(* IEC 61131-3 sources: plc-process-lib/tests/POUs/Suites/FB_Pid_Test, 85 files *)

(* ---- AntiWindupLongSaturationRecoversWithinTt.method.decl.st ---- *)
// Anti-windup обратным расчётом (Kp = 1, Ti = 10 с, Tt = авто = Ti): 60 с на верхнем пределе при
// ошибке +20 %, затем ошибка -20 %. С обратным расчётом интегратор ограничен (v ≈ 100 + Tt·Kp·e/Ti)
// и выход уходит с предела сразу; для сравнения тот же ФБ с Tt = 1·10^6 с (обратного расчёта
// практически нет) остаётся на пределе и через Tt после смены знака.
METHOD PRIVATE AntiWindupLongSaturationRecoversWithinTt
VAR
    fbTime    : FB_FakeTime;       // подменное время, старт 1 ч
    fbPidAw   : FB_PID;            // ФБ под тестом: Tt = авто
    fbPidNoAw : FB_PID;            // сравнение: Tt = 1e6 с
    stCmdAw   : ST_PidCmd;         // команды
    stCmdNoAw : ST_PidCmd;
    stRetAw   : ST_DeviceRetain;   // режим: старт в Manual
    stRetNoAw : ST_DeviceRetain;
    stCfgAw   : ST_PidCfg;         // конфигурация
    stCfgNoAw : ST_PidCfg;
    iStep     : INT;               // шаг цикла
    rOutSatAw : REAL;              // выход в конце насыщения
    rISatAw   : REAL;              // интегратор в конце насыщения
    rISatNoAw : REAL;
    rOutRevAw : REAL;              // выход в первом шаге после смены знака ошибки
    rOutRevNo : REAL;
END_VAR

(* ---- AntiWindupLongSaturationRecoversWithinTt.method.impl.st ---- *)
coUnit.TEST('Pid_AntiWindup_LongSaturation_RecoversWithinTt');
// источник: tools/reference/pid.py, сценарий aw_recovery
stCfgAw.rKp := 1.0;
stCfgAw.rTi_s := 10.0;
stCfgAw.rTt_s := 0.0;
stCfgNoAw := stCfgAw;
stCfgNoAw.rTt_s := 1.0E6;
stCmdAw.rManualOut_pct := 50.0;
stCmdAw.rSp_eu := 50.0;
stCmdNoAw := stCmdAw;
fbPidAw.rPv_eu := 50.0;
fbPidAw.xPvValid := TRUE;
fbPidNoAw.rPv_eu := 50.0;
fbPidNoAw.xPvValid := TRUE;
fbPidAw(itfTime := fbTime, stCmd := stCmdAw, stRetain := stRetAw, stCfg := stCfgAw);          // t0: Manual
fbPidNoAw(itfTime := fbTime, stCmd := stCmdNoAw, stRetain := stRetNoAw, stCfg := stCfgNoAw);
fbTime.Advance(tStep := T#100MS);
stCmdAw.stCommon.xSetAuto := TRUE;
stCmdNoAw.stCommon.xSetAuto := TRUE;
fbPidAw(itfTime := fbTime, stCmd := stCmdAw, stRetain := stRetAw, stCfg := stCfgAw);          // Auto
fbPidNoAw(itfTime := fbTime, stCmd := stCmdNoAw, stRetain := stRetNoAw, stCfg := stCfgNoAw);
fbPidAw.rPv_eu := 30.0;                                                                         // e = +20 %
fbPidNoAw.rPv_eu := 30.0;
FOR iStep := 1 TO 600 DO                                                                        // 60 с
    fbTime.Advance(tStep := T#100MS);
    fbPidAw(itfTime := fbTime, stCmd := stCmdAw, stRetain := stRetAw, stCfg := stCfgAw);
    fbPidNoAw(itfTime := fbTime, stCmd := stCmdNoAw, stRetain := stRetNoAw, stCfg := stCfgNoAw);
END_FOR
rOutSatAw := fbPidAw.rOut_pct;
rISatAw := fbPidAw.stSts.rI_pct;
rISatNoAw := fbPidNoAw.stSts.rI_pct;
fbPidAw.rPv_eu := 70.0;                                                                         // e = -20 %
fbPidNoAw.rPv_eu := 70.0;
fbTime.Advance(tStep := T#100MS);
fbPidAw(itfTime := fbTime, stCmd := stCmdAw, stRetain := stRetAw, stCfg := stCfgAw);
fbPidNoAw(itfTime := fbTime, stCmd := stCmdNoAw, stRetain := stRetNoAw, stCfg := stCfgNoAw);
rOutRevAw := fbPidAw.rOut_pct;
rOutRevNo := fbPidNoAw.rOut_pct;
FOR iStep := 1 TO 99 DO                                                                         // до Tt = 10 с
    fbTime.Advance(tStep := T#100MS);
    fbPidAw(itfTime := fbTime, stCmd := stCmdAw, stRetain := stRetAw, stCfg := stCfgAw);
    fbPidNoAw(itfTime := fbTime, stCmd := stCmdNoAw, stRetain := stRetNoAw, stCfg := stCfgNoAw);
END_FOR
// ref: aw_recovery.out_sat_aw
AssertEquals_REAL(Expected := 100.0, Actual := rOutSatAw, Delta := 1.0E-4, Message := 'saturated at rOutMax_pct');
// ref: aw_recovery.i_sat_aw
AssertEquals_REAL(Expected := 99.782799, Actual := rISatAw, Delta := 1.0E-3,
                  Message := 'I bounded by back-calculation');
// ref: aw_recovery.i_sat_noaw
AssertEquals_REAL(Expected := 169.997986, Actual := rISatNoAw, Delta := 1.0E-3, Message := 'I winds up without it');
// ref: aw_recovery.out_rev_aw
AssertEquals_REAL(Expected := 79.782799, Actual := rOutRevAw, Delta := 1.0E-3, Message := 'leaves limit at once');
// ref: aw_recovery.out_rev_noaw
AssertEquals_REAL(Expected := 100.0, Actual := rOutRevNo, Delta := 1.0E-4, Message := 'wound-up: still at limit');
// ref: aw_recovery.out_tt_aw
AssertEquals_REAL(Expected := 59.982796, Actual := fbPidAw.rOut_pct, Delta := 1.0E-3, Message := 'recovered within Tt');
// ref: aw_recovery.out_tt_noaw
AssertEquals_REAL(Expected := 100.0, Actual := fbPidNoAw.rOut_pct, Delta := 1.0E-4, Message := 'wound-up after Tt');
AssertFalse(Condition := fbPidAw.xSatHigh, Message := 'back-calculation: not saturated after Tt');
coUnit.TEST_FINISHED();

(* ---- AntiWindupOutActFeedbackTracksExternalLimit.method.decl.st ---- *)
// Обратный расчёт по фактическому выходу (xUseOutAct): механизм не опускается ниже 30 % (минимум
// частоты ПЧ), rOutAct_pct = MAX(30, выход прошлого вызова). При ошибке -10 % 60 с выход ПИД
// держится у внешнего предела (около 30 - Tt·Kp·|e|/Ti = 20 %), а не уходит в 0; после смены
// знака ошибки механизм отвечает сразу. Без xUseOutAct ПИД уходит в 0 и после смены знака
// остаётся ниже 30 %.
METHOD PRIVATE AntiWindupOutActFeedbackTracksExternalLimit
VAR
    fbTime     : FB_FakeTime;       // подменное время, старт 1 ч
    fbPidAct   : FB_PID;            // ФБ под тестом: xUseOutAct
    fbPidNoAct : FB_PID;            // сравнение: без xUseOutAct
    stCmdAct   : ST_PidCmd;         // команды
    stCmdNoAct : ST_PidCmd;
    stRetAct   : ST_DeviceRetain;   // режим: старт в Manual
    stRetNoAct : ST_DeviceRetain;
    stCfgAct   : ST_PidCfg;         // конфигурация
    stCfgNoAct : ST_PidCfg;
    iStep      : INT;               // шаг цикла
    rHoldAct   : REAL;              // выход в конце 60 с
    rHoldNoAct : REAL;
END_VAR

(* ---- AntiWindupOutActFeedbackTracksExternalLimit.method.impl.st ---- *)
coUnit.TEST('Pid_AntiWindup_OutActFeedback_TracksExternalLimit');
// источник: tools/reference/pid.py, сценарий outact
stCfgAct.rKp := 1.0;
stCfgAct.rTi_s := 10.0;
stCfgNoAct := stCfgAct;
stCfgAct.xUseOutAct := TRUE;
stCmdAct.rManualOut_pct := 50.0;
stCmdAct.rSp_eu := 50.0;
stCmdNoAct := stCmdAct;
fbPidAct.rPv_eu := 50.0;
fbPidAct.xPvValid := TRUE;
fbPidNoAct.rPv_eu := 50.0;
fbPidNoAct.xPvValid := TRUE;
fbPidAct(itfTime := fbTime, stCmd := stCmdAct, stRetain := stRetAct, stCfg := stCfgAct);          // t0: Manual
fbPidNoAct(itfTime := fbTime, stCmd := stCmdNoAct, stRetain := stRetNoAct, stCfg := stCfgNoAct);
fbPidAct.rOutAct_pct := MAX(30.0, fbPidAct.rOut_pct);
fbPidNoAct.rOutAct_pct := MAX(30.0, fbPidNoAct.rOut_pct);
fbTime.Advance(tStep := T#100MS);
stCmdAct.stCommon.xSetAuto := TRUE;
stCmdNoAct.stCommon.xSetAuto := TRUE;
fbPidAct(itfTime := fbTime, stCmd := stCmdAct, stRetain := stRetAct, stCfg := stCfgAct);          // Auto
fbPidNoAct(itfTime := fbTime, stCmd := stCmdNoAct, stRetain := stRetNoAct, stCfg := stCfgNoAct);
fbPidAct.rPv_eu := 60.0;                                                                            // e = -10 %
fbPidNoAct.rPv_eu := 60.0;
FOR iStep := 1 TO 600 DO                                                                            // 60 с
    fbPidAct.rOutAct_pct := MAX(30.0, fbPidAct.rOut_pct);
    fbPidNoAct.rOutAct_pct := MAX(30.0, fbPidNoAct.rOut_pct);
    fbTime.Advance(tStep := T#100MS);
    fbPidAct(itfTime := fbTime, stCmd := stCmdAct, stRetain := stRetAct, stCfg := stCfgAct);
    fbPidNoAct(itfTime := fbTime, stCmd := stCmdNoAct, stRetain := stRetNoAct, stCfg := stCfgNoAct);
END_FOR
rHoldAct := fbPidAct.rOut_pct;
rHoldNoAct := fbPidNoAct.rOut_pct;
fbPidAct.rPv_eu := 40.0;                                                                            // e = +10 %
fbPidNoAct.rPv_eu := 40.0;
FOR iStep := 1 TO 30 DO                                                                             // 3 с
    fbPidAct.rOutAct_pct := MAX(30.0, fbPidAct.rOut_pct);
    fbPidNoAct.rOutAct_pct := MAX(30.0, fbPidNoAct.rOut_pct);
    fbTime.Advance(tStep := T#100MS);
    fbPidAct(itfTime := fbTime, stCmd := stCmdAct, stRetain := stRetAct, stCfg := stCfgAct);
    fbPidNoAct(itfTime := fbTime, stCmd := stCmdNoAct, stRetain := stRetNoAct, stCfg := stCfgNoAct);
END_FOR
// ref: outact.out_hold_act
AssertEquals_REAL(Expected := 20.067717, Actual := rHoldAct, Delta := 1.0E-3, Message := 'held near external limit');
// ref: outact.out_hold_noact
AssertEquals_REAL(Expected := 0.0, Actual := rHoldNoAct, Delta := 1.0E-4, Message := 'without OutAct: down to 0');
// ref: outact.out_rev_act
AssertEquals_REAL(Expected := 42.839634, Actual := fbPidAct.rOut_pct, Delta := 1.0E-3, Message := 'responds at once');
// ref: outact.out_rev_noact
AssertEquals_REAL(Expected := 14.239797, Actual := fbPidNoAct.rOut_pct, Delta := 1.0E-3, Message := 'still below 30 %');
AssertTrue(Condition := fbPidAct.rOut_pct > 30.0, Message := 'with OutAct the actuator moves above its minimum');
AssertTrue(Condition := fbPidNoAct.rOut_pct < 30.0, Message := 'without OutAct the actuator still sits at 30 %');
coUnit.TEST_FINISHED();

(* ---- AntiWindupOutActNaNUsesOwnOutput.method.decl.st ---- *)
// xUseOutAct, а фактический выход не конечен (связь с ПЧ потеряна, в образе обмена NaN): обратный
// расчёт идёт по собственному выходу ФБ, NaN в интегратор не попадает. Без насыщения член u - v
// равен нулю — выход тот же, что в сценарии integral.
METHOD PRIVATE AntiWindupOutActNaNUsesOwnOutput
VAR
    fbTime   : FB_FakeTime;       // подменное время, старт 1 ч
    fbPid    : FB_PID;            // ФБ под тестом
    stCmd    : ST_PidCmd;         // команды
    stRetain : ST_DeviceRetain;   // режим
    stCfg    : ST_PidCfg;         // конфигурация теста
    uBits    : U_RealBits;        // источник NaN
    iStep    : INT;               // шаг цикла
    rOut1    : REAL;              // выход первого шага в Auto
END_VAR

(* ---- AntiWindupOutActNaNUsesOwnOutput.method.impl.st ---- *)
coUnit.TEST('Pid_AntiWindup_OutActNaN_UsesOwnOutput');
// источник: tools/reference/pid.py, сценарий outact_nan
uBits.dwValue := 16#7FC00000;                                                          // тихий NaN
stCfg.rKp := 2.0;
stCfg.rTi_s := 10.0;
stCfg.xUseOutAct := TRUE;
stCmd.rManualOut_pct := 30.0;
stCmd.rSp_eu := 50.0;
fbPid.rPv_eu := 50.0;
fbPid.xPvValid := TRUE;
fbPid.rOutAct_pct := uBits.rValue;                                                     // фактический выход неизвестен
fbPid(itfTime := fbTime, stCmd := stCmd, stRetain := stRetain, stCfg := stCfg);       // t0: Manual
fbTime.Advance(tStep := T#100MS);
stCmd.stCommon.xSetAuto := TRUE;
fbPid(itfTime := fbTime, stCmd := stCmd, stRetain := stRetain, stCfg := stCfg);       // Auto
fbPid.rPv_eu := 46.0;                                                                  // e = 4 %
fbTime.Advance(tStep := T#100MS);
fbPid(itfTime := fbTime, stCmd := stCmd, stRetain := stRetain, stCfg := stCfg);
rOut1 := fbPid.rOut_pct;
FOR iStep := 1 TO 50 DO
    fbTime.Advance(tStep := T#100MS);
    fbPid(itfTime := fbTime, stCmd := stCmd, stRetain := stRetain, stCfg := stCfg);
END_FOR
// AssertEquals_REAL пропускает NaN (ABS(NaN) > Delta = FALSE): конечность проверяется отдельно
AssertTrue(Condition := F_IsFinite(rIn := fbPid.stSts.rI_pct), Message := 'integrator stays finite');
AssertTrue(Condition := F_IsFinite(rIn := fbPid.rOut_pct), Message := 'output stays finite');
// ref: outact_nan.out_first
AssertEquals_REAL(Expected := 38.0, Actual := rOut1, Delta := 1.0E-4, Message := 'first step: 30 + P');
// ref: outact_nan.out_after_5s
AssertEquals_REAL(Expected := 42.0, Actual := fbPid.rOut_pct, Delta := 1.0E-4, Message := 'integral as usual');
// ref: outact_nan.i_after_5s
AssertEquals_REAL(Expected := 34.080002, Actual := fbPid.stSts.rI_pct, Delta := 1.0E-4, Message := 'integrator finite');
coUnit.TEST_FINISHED();

(* ---- AntiWindupTtBelowDtGainClampedToOne.method.decl.st ---- *)
// Постоянная слежения меньше шага (Tt = 0,05 с, dt = 0,1 с): множитель обратного расчёта
// MIN(dt/Tt, 1) = 1, и за один шаг насыщения интегратор садится ровно на v = u (I = 1 %), выход
// остаётся на пределе. Без MIN множитель был бы 2: I = -49 %, и на следующем шаге выход упал бы с
// предела до 51 % при той же ошибке +50 % — колебание обратного расчёта.
METHOD PRIVATE AntiWindupTtBelowDtGainClampedToOne
VAR
    fbTime   : FB_FakeTime;       // подменное время, старт 1 ч
    fbPid    : FB_PID;            // ФБ под тестом
    stCmd    : ST_PidCmd;         // команды
    stRetain : ST_DeviceRetain;   // режим: старт в Manual
    stCfg    : ST_PidCfg;         // конфигурация теста
    iStep    : INT;               // шаг цикла
    rOutSat  : REAL;              // выход в первом шаге насыщения
    rISat    : REAL;              // интегратор в первом шаге насыщения
    rOutNext : REAL;              // выход в следующем шаге
    rINext   : REAL;              // интегратор в следующем шаге
END_VAR

(* ---- AntiWindupTtBelowDtGainClampedToOne.method.impl.st ---- *)
coUnit.TEST('Pid_AntiWindup_TtBelowDt_GainClampedToOne');
// источник: tools/reference/pid.py, сценарий tt_small
stCfg.rKp := 2.0;
stCfg.rTi_s := 10.0;
stCfg.rTt_s := 0.05;                                                                   // Tt < dt
stCmd.rManualOut_pct := 50.0;
stCmd.rSp_eu := 50.0;
fbPid.rPv_eu := 50.0;
fbPid.xPvValid := TRUE;
fbPid(itfTime := fbTime, stCmd := stCmd, stRetain := stRetain, stCfg := stCfg);       // t0: Manual
fbTime.Advance(tStep := T#100MS);
stCmd.stCommon.xSetAuto := TRUE;
fbPid(itfTime := fbTime, stCmd := stCmd, stRetain := stRetain, stCfg := stCfg);       // Auto, I = 50 %
fbPid.rPv_eu := 0.0;                                                                   // e = +50 %, v = 150 %
fbTime.Advance(tStep := T#100MS);
fbPid(itfTime := fbTime, stCmd := stCmd, stRetain := stRetain, stCfg := stCfg);
rOutSat := fbPid.rOut_pct;
rISat := fbPid.stSts.rI_pct;
fbTime.Advance(tStep := T#100MS);
fbPid(itfTime := fbTime, stCmd := stCmd, stRetain := stRetain, stCfg := stCfg);
rOutNext := fbPid.rOut_pct;
rINext := fbPid.stSts.rI_pct;
FOR iStep := 1 TO 8 DO                                                                 // до 1 с насыщения
    fbTime.Advance(tStep := T#100MS);
    fbPid(itfTime := fbTime, stCmd := stCmd, stRetain := stRetain, stCfg := stCfg);
END_FOR
// ref: tt_small.out_sat
AssertEquals_REAL(Expected := 100.0, Actual := rOutSat, Delta := 1.0E-4, Message := 'saturated at rOutMax_pct');
// ref: tt_small.i_sat
AssertEquals_REAL(Expected := 1.0, Actual := rISat, Delta := 1.0E-4,
                  Message := 'gain clamped to 1: I = 50 + 1 - 50, not -49');
// ref: tt_small.out_next
AssertEquals_REAL(Expected := 100.0, Actual := rOutNext, Delta := 1.0E-4,
                  Message := 'next step stays at limit (no back-calculation oscillation)');
// ref: tt_small.i_next
AssertEquals_REAL(Expected := 1.0, Actual := rINext, Delta := 1.0E-4, Message := 'I settles at v = u');
// ref: tt_small.out_1s
AssertEquals_REAL(Expected := 100.0, Actual := fbPid.rOut_pct, Delta := 1.0E-4, Message := 'at limit after 1 s');
AssertTrue(Condition := fbPid.xSatHigh, Message := 'xSatHigh while saturated');
coUnit.TEST_FINISHED();

(* ---- CfgChecksSetDocumentedBits.method.decl.st ---- *)
// CheckConfig: каждая неверная группа параметров даёт свой бит wCfgErr (карта битов
// docs/fb/FB_PID.md); значения вне строгих перечислений — через объединение U_TestPidEnumInt,
// NaN — через U_RealBits.
METHOD PRIVATE CfgChecksSetDocumentedBits
VAR
    fbTime   : FB_FakeTime;        // подменное время, старт 1 ч
    fbPid    : FB_PID;             // ФБ под тестом
    stCmd    : ST_PidCmd;          // команды
    stRetain : ST_DeviceRetain;    // режим: Manual
    stCfgDef : ST_PidCfg;          // конфигурация по умолчанию
    stCfg    : ST_PidCfg;          // проверяемая конфигурация
    stSlot   : ST_AlarmCfg;        // копия слота тревоги
    uBad     : U_TestPidEnumInt;   // значение вне перечислений
    uBits    : U_RealBits;         // источник NaN
END_VAR

(* ---- CfgSpLimitsEqualFixedSetpoint.method.decl.st ---- *)
// Равные пределы задания допустимы (бит 6 — только min > max): задание фиксировано, любое
// задание оператора ограничивается этим значением.
METHOD PRIVATE CfgSpLimitsEqualFixedSetpoint
VAR
    fbTime   : FB_FakeTime;       // подменное время, старт 1 ч
    fbPid    : FB_PID;            // ФБ под тестом
    stCmd    : ST_PidCmd;         // команды
    stRetain : ST_DeviceRetain;   // режим
    stCfg    : ST_PidCfg;         // конфигурация теста
END_VAR

(* ---- DeadbandNoActionInsideBand.method.decl.st ---- *)
// Зона нечувствительности 1 % (Kp = 2, Ti = 10 с): ошибка 0,8 % — e' = 0, выход и интегратор
// стоят 2 с, бит IN_DEADBAND; ошибка 1,5 % — e' = 0,5 %, выход +1 % без скачка на границе зоны.
METHOD PRIVATE DeadbandNoActionInsideBand
VAR
    fbTime   : FB_FakeTime;       // подменное время, старт 1 ч
    fbPid    : FB_PID;            // ФБ под тестом
    stCmd    : ST_PidCmd;         // команды
    stRetain : ST_DeviceRetain;   // режим: старт в Manual
    stCfg    : ST_PidCfg;         // конфигурация теста
    iStep    : INT;               // шаг цикла
    rOutIn   : REAL;              // выход в зоне
    rErrIn   : REAL;              // e' в зоне
    wStsIn   : WORD;              // wStatus в зоне
END_VAR

(* ---- DeadbandNoActionInsideBand.method.impl.st ---- *)
coUnit.TEST('Pid_Deadband_NoActionInsideBand');
// источник: tools/reference/pid.py, сценарий deadband
stCfg.rKp := 2.0;
stCfg.rTi_s := 10.0;
stCfg.rDeadband_pct := 1.0;
stCmd.rManualOut_pct := 30.0;
stCmd.rSp_eu := 50.0;
fbPid.rPv_eu := 50.0;
fbPid.xPvValid := TRUE;
fbPid(itfTime := fbTime, stCmd := stCmd, stRetain := stRetain, stCfg := stCfg);       // t0: Manual
fbTime.Advance(tStep := T#100MS);
stCmd.stCommon.xSetAuto := TRUE;
fbPid(itfTime := fbTime, stCmd := stCmd, stRetain := stRetain, stCfg := stCfg);       // Auto
fbPid.rPv_eu := 49.2;                                                                  // e = 0,8 %
FOR iStep := 1 TO 20 DO
    fbTime.Advance(tStep := T#100MS);
    fbPid(itfTime := fbTime, stCmd := stCmd, stRetain := stRetain, stCfg := stCfg);
END_FOR
rOutIn := fbPid.rOut_pct;
rErrIn := fbPid.stSts.rErr_pct;
wStsIn := fbPid.stSts.stCommon.wStatus;
fbPid.rPv_eu := 48.5;                                                                  // e = 1,5 %
fbTime.Advance(tStep := T#100MS);
fbPid(itfTime := fbTime, stCmd := stCmd, stRetain := stRetain, stCfg := stCfg);
// ref: deadband.out_inside
AssertEquals_REAL(Expected := 30.0, Actual := rOutIn, Delta := 1.0E-4, Message := 'no action inside band');
// ref: deadband.err_inside
AssertEquals_REAL(Expected := 0.0, Actual := rErrIn, Delta := 1.0E-6, Message := 'e prime = 0 inside band');
AssertEquals_WORD(Expected := GVL_Const.PID_STS_IN_DEADBAND, Actual := wStsIn AND GVL_Const.PID_STS_IN_DEADBAND,
                  Message := 'status bit IN_DEADBAND');
// ref: deadband.out_outside
AssertEquals_REAL(Expected := 31.0, Actual := fbPid.rOut_pct, Delta := 1.0E-4, Message := 'out = 30 + 2 * (1.5 - 1)');
// ref: deadband.err_outside
AssertEquals_REAL(Expected := 0.5, Actual := fbPid.stSts.rErr_pct, Delta := 1.0E-4, Message := 'e prime = e - band');
AssertEquals_WORD(Expected := 0, Actual := fbPid.stSts.stCommon.wStatus AND GVL_Const.PID_STS_IN_DEADBAND,
                  Message := 'IN_DEADBAND cleared');
coUnit.TEST_FINISHED();

(* ---- DefaultCfgPassesCheck.method.decl.st ---- *)
// Значения ST_PidCfg по умолчанию проходят CheckConfig (инвариант генератора iolistgen, контракт
// 2.3): wCfgErr = 0, бита CFG_ERROR нет, статус Good в Manual.
METHOD PRIVATE DefaultCfgPassesCheck
VAR
    fbTime   : FB_FakeTime;       // подменное время, старт 1 ч
    fbPid    : FB_PID;            // ФБ под тестом
    stCmd    : ST_PidCmd;         // команды
    stRetain : ST_DeviceRetain;   // режим: Manual
    stCfg    : ST_PidCfg;         // конфигурация по умолчанию
END_VAR

(* ---- DFilterPvStepDecaysWithTdOverN.method.decl.st ---- *)
// Фильтр Д (Td = 5 с, N = 10, Tf = 0,5 с, шаг 100 мс): после ступени PV составляющая D затухает
// множителем Tf/(Tf + dt) за шаг; через Tf от неё остаётся (5/6)^5, около 0,40.
METHOD PRIVATE DFilterPvStepDecaysWithTdOverN
VAR
    fbTime   : FB_FakeTime;       // подменное время, старт 1 ч
    fbPid    : FB_PID;            // ФБ под тестом
    stCmd    : ST_PidCmd;         // команды
    stRetain : ST_DeviceRetain;   // режим: старт в Manual
    stCfg    : ST_PidCfg;         // конфигурация теста
    iStep    : INT;               // шаг цикла
    rD1      : REAL;              // D сразу после ступени
END_VAR

(* ---- DFilterPvStepDecaysWithTdOverN.method.impl.st ---- *)
coUnit.TEST('Pid_DFilter_PvStep_DecaysWithTdOverN');
// источник: tools/reference/pid.py, сценарий d_filter
stCfg.rKp := 1.0;
stCfg.rTi_s := 0.0;
stCfg.rTd_s := 5.0;
stCfg.rDFilterN := 10.0;
stCmd.rManualOut_pct := 50.0;
stCmd.rSp_eu := 50.0;
fbPid.rPv_eu := 50.0;
fbPid.xPvValid := TRUE;
fbPid(itfTime := fbTime, stCmd := stCmd, stRetain := stRetain, stCfg := stCfg);       // t0: Manual
fbTime.Advance(tStep := T#100MS);
stCmd.stCommon.xSetAuto := TRUE;
fbPid(itfTime := fbTime, stCmd := stCmd, stRetain := stRetain, stCfg := stCfg);       // Auto
fbPid.rPv_eu := 52.0;                                                                  // ступень PV
fbTime.Advance(tStep := T#100MS);
fbPid(itfTime := fbTime, stCmd := stCmd, stRetain := stRetain, stCfg := stCfg);
rD1 := fbPid.stSts.rD_pct;
FOR iStep := 1 TO 5 DO                                                                 // ещё Tf = 0,5 с
    fbTime.Advance(tStep := T#100MS);
    fbPid(itfTime := fbTime, stCmd := stCmd, stRetain := stRetain, stCfg := stCfg);
END_FOR
// ref: d_filter.d_step
AssertEquals_REAL(Expected := -16.666666, Actual := rD1, Delta := 1.0E-4, Message := 'D right after PV step');
// ref: d_filter.d_after_tf
AssertEquals_REAL(Expected := -6.697959, Actual := fbPid.stSts.rD_pct, Delta := 1.0E-4, Message := 'D after Tf');
// ref: d_filter.ratio
AssertEquals_REAL(Expected := 0.401878, Actual := fbPid.stSts.rD_pct / rD1, Delta := 1.0E-5,
                  Message := 'decay (Tf / (Tf + dt))^5 over Tf = Td / N');
coUnit.TEST_FINISHED();

(* ---- DirectActionInvertsSign.method.decl.st ---- *)
// Прямое и обратное действие (Kp = 2, без I): при PV на 10 % выше задания обратное действие
// уменьшает выход на 20 %, прямое — увеличивает; знак ошибки в Sts — со знаком действия.
METHOD PRIVATE DirectActionInvertsSign
VAR
    fbTime   : FB_FakeTime;       // подменное время, старт 1 ч
    fbPidRev : FB_PID;            // обратное действие
    fbPidDir : FB_PID;            // прямое действие
    stCmdRev : ST_PidCmd;         // команды
    stCmdDir : ST_PidCmd;
    stRetRev : ST_DeviceRetain;   // режим: старт в Manual
    stRetDir : ST_DeviceRetain;
    stCfgRev : ST_PidCfg;         // конфигурация
    stCfgDir : ST_PidCfg;
END_VAR

(* ---- DOnMeasurementSetpointStepNoDerivativeKick.method.decl.st ---- *)
// D по измерению (Kp = 1, Td = 5 с, N = 10, без I): ступень задания меняет выход только на P
// (D = 0, «удара» нет), ступень PV на 2 % даёт D = -Kp·Td/(Tf + dt)·2 %.
METHOD PRIVATE DOnMeasurementSetpointStepNoDerivativeKick
VAR
    fbTime   : FB_FakeTime;       // подменное время, старт 1 ч
    fbPid    : FB_PID;            // ФБ под тестом
    stCmd    : ST_PidCmd;         // команды
    stRetain : ST_DeviceRetain;   // режим: старт в Manual
    stCfg    : ST_PidCfg;         // конфигурация теста
END_VAR

(* ---- DtGapBoundaryAtTDtMax.method.decl.st ---- *)
// Граница разрыва времени (tDtMax = 1 с): шаг ровно 1 с — обычный расчёт (dt = 1000 мс, интеграл
// +0,8 %, без DT_GAP), шаг 1,001 с — разрыв: шаг инициализации, выход прежний, интегратор
// предустановлен I := u - P (30,8 %), бит DT_GAP. Условие контракта — «dt > tDtMax».
METHOD PRIVATE DtGapBoundaryAtTDtMax
VAR
    fbTime   : FB_FakeTime;       // подменное время, старт 1 ч
    fbPid    : FB_PID;            // ФБ под тестом
    stCmd    : ST_PidCmd;         // команды
    stRetain : ST_DeviceRetain;   // режим: старт в Manual
    stCfg    : ST_PidCfg;         // конфигурация теста
    iStep    : INT;               // шаг цикла
    rIBefore : REAL;              // интегратор до длинных шагов
    rIAtMax  : REAL;              // интегратор после шага ровно tDtMax
    rDtAtMax : REAL;              // stSts.rDt_ms после шага ровно tDtMax
    wStsMax  : WORD;              // wStatus после шага ровно tDtMax
    rOutMax  : REAL;              // выход после шага ровно tDtMax
END_VAR

(* ---- DtGapBoundaryAtTDtMax.method.impl.st ---- *)
coUnit.TEST('Pid_DtGap_BoundaryAtTDtMax');
// источник: tools/reference/pid.py, сценарий dt_boundary
stCfg.rKp := 2.0;
stCfg.rTi_s := 10.0;
stCfg.tDtMax := T#1S;
stCmd.rManualOut_pct := 30.0;
stCmd.rSp_eu := 50.0;
fbPid.rPv_eu := 50.0;
fbPid.xPvValid := TRUE;
fbPid(itfTime := fbTime, stCmd := stCmd, stRetain := stRetain, stCfg := stCfg);       // t0: Manual
fbTime.Advance(tStep := T#100MS);
stCmd.stCommon.xSetAuto := TRUE;
fbPid(itfTime := fbTime, stCmd := stCmd, stRetain := stRetain, stCfg := stCfg);       // Auto
fbPid.rPv_eu := 46.0;                                                                  // e = 4 %
FOR iStep := 1 TO 10 DO
    fbTime.Advance(tStep := T#100MS);
    fbPid(itfTime := fbTime, stCmd := stCmd, stRetain := stRetain, stCfg := stCfg);
END_FOR
rIBefore := fbPid.stSts.rI_pct;
fbTime.Advance(tStep := T#1S);                                                         // ровно tDtMax
fbPid(itfTime := fbTime, stCmd := stCmd, stRetain := stRetain, stCfg := stCfg);
rIAtMax := fbPid.stSts.rI_pct;
rDtAtMax := fbPid.stSts.rDt_ms;
wStsMax := fbPid.stSts.stCommon.wStatus;
rOutMax := fbPid.rOut_pct;
fbTime.Advance(tStep := T#1001MS);                                                     // на 1 мс больше
fbPid(itfTime := fbTime, stCmd := stCmd, stRetain := stRetain, stCfg := stCfg);
// ref: dt_boundary.i_before
AssertEquals_REAL(Expected := 30.8, Actual := rIBefore, Delta := 1.0E-4, Message := 'I before long steps');
// ref: dt_boundary.i_at_max
AssertEquals_REAL(Expected := 31.6, Actual := rIAtMax, Delta := 1.0E-4, Message := 'dt = tDtMax integrated (+0.8)');
// ref: dt_boundary.dt_ms_at_max
AssertEquals_REAL(Expected := 1000.0, Actual := rDtAtMax, Delta := 1.0E-3, Message := 'rDt_ms = 1000 at tDtMax');
AssertEquals_WORD(Expected := 0, Actual := wStsMax AND GVL_Const.PID_STS_DT_GAP, Message := 'no DT_GAP at tDtMax');
// ref: dt_boundary.i_over_max
AssertEquals_REAL(Expected := 30.8, Actual := fbPid.stSts.rI_pct, Delta := 1.0E-4,
                  Message := 'dt > tDtMax: init step presets I = u - P');
// ref: dt_boundary.out_over_max
AssertEquals_REAL(Expected := 38.8, Actual := fbPid.rOut_pct, Delta := 1.0E-4, Message := 'gap: output held');
AssertEquals_REAL(Expected := rOutMax, Actual := fbPid.rOut_pct, Delta := 0.0,
                  Message := 'gap: exactly previous output');
AssertEquals_WORD(Expected := GVL_Const.PID_STS_DT_GAP,
                  Actual := fbPid.stSts.stCommon.wStatus AND GVL_Const.PID_STS_DT_GAP,
                  Message := 'DT_GAP above tDtMax');
AssertEquals_REAL(Expected := 0.0, Actual := fbPid.stSts.rDt_ms, Delta := 0.0, Message := 'rDt_ms = 0 on init step');
coUnit.TEST_FINISHED();

(* ---- DtGapSkipsIntegration.method.decl.st ---- *)
// Разрыв времени 5 с > tDtMax = 2 с (стоп ПЛК, отладка): шаг инициализации — выход прежний,
// интегратор не получает 5 с (без защиты было бы +4 %), бит DT_GAP и предупреждение
// PID_WRN_DT_GAP на один вызов; дальше интегрирование по обычному шагу.
METHOD PRIVATE DtGapSkipsIntegration
VAR
    fbTime    : FB_FakeTime;       // подменное время, старт 1 ч
    fbPid     : FB_PID;            // ФБ под тестом
    stCmd     : ST_PidCmd;         // команды
    stRetain  : ST_DeviceRetain;   // режим: старт в Manual
    stCfg     : ST_PidCfg;         // конфигурация теста
    iStep     : INT;               // шаг цикла
    rBefore   : REAL;              // выход до разрыва
    rGap      : REAL;              // выход в вызове после разрыва
    wStsGap   : WORD;              // wStatus в вызове после разрыва
    wWrnGap   : WORD;              // wWarning в вызове после разрыва
    rAfter    : REAL;              // выход в следующем вызове
    wStsAfter : WORD;              // wStatus в следующем вызове
END_VAR

(* ---- DtGapSkipsIntegration.method.impl.st ---- *)
coUnit.TEST('Pid_DtGap_SkipsIntegration');
// источник: tools/reference/pid.py, сценарий dt_gap
stCfg.rKp := 2.0;
stCfg.rTi_s := 10.0;
stCmd.rManualOut_pct := 30.0;
stCmd.rSp_eu := 50.0;
fbPid.rPv_eu := 50.0;
fbPid.xPvValid := TRUE;
fbPid(itfTime := fbTime, stCmd := stCmd, stRetain := stRetain, stCfg := stCfg);       // t0: Manual
fbTime.Advance(tStep := T#100MS);
stCmd.stCommon.xSetAuto := TRUE;
fbPid(itfTime := fbTime, stCmd := stCmd, stRetain := stRetain, stCfg := stCfg);       // Auto
fbPid.rPv_eu := 46.0;                                                                  // e = 4 %
FOR iStep := 1 TO 10 DO
    fbTime.Advance(tStep := T#100MS);
    fbPid(itfTime := fbTime, stCmd := stCmd, stRetain := stRetain, stCfg := stCfg);
END_FOR
rBefore := fbPid.rOut_pct;
fbTime.Advance(tStep := T#5S);                                                         // разрыв
fbPid(itfTime := fbTime, stCmd := stCmd, stRetain := stRetain, stCfg := stCfg);
rGap := fbPid.rOut_pct;
wStsGap := fbPid.stSts.stCommon.wStatus;
wWrnGap := fbPid.stSts.stCommon.wWarning;
fbTime.Advance(tStep := T#100MS);
fbPid(itfTime := fbTime, stCmd := stCmd, stRetain := stRetain, stCfg := stCfg);
rAfter := fbPid.rOut_pct;
wStsAfter := fbPid.stSts.stCommon.wStatus;
fbTime.Advance(tStep := T#100MS);
fbPid(itfTime := fbTime, stCmd := stCmd, stRetain := stRetain, stCfg := stCfg);
// ref: dt_gap.out_before
AssertEquals_REAL(Expected := 38.72, Actual := rBefore, Delta := 1.0E-4, Message := 'output before gap');
// ref: dt_gap.out_gap
AssertEquals_REAL(Expected := 38.72, Actual := rGap, Delta := 1.0E-4,
                  Message := 'gap: output held, no 5 s integration');
AssertEquals_WORD(Expected := GVL_Const.PID_STS_DT_GAP, Actual := wStsGap AND GVL_Const.PID_STS_DT_GAP,
                  Message := 'status bit DT_GAP on gap');
AssertEquals_WORD(Expected := GVL_Const.PID_WRN_DT_GAP, Actual := wWrnGap, Message := 'warning DT_GAP on gap');
// ref: dt_gap.out_after
AssertEquals_REAL(Expected := 38.72, Actual := rAfter, Delta := 1.0E-4, Message := 'first normal step after gap');
AssertEquals_WORD(Expected := 0, Actual := wStsAfter AND GVL_Const.PID_STS_DT_GAP, Message := 'DT_GAP for one call');
// ref: dt_gap.out_after2
AssertEquals_REAL(Expected := 38.8, Actual := fbPid.rOut_pct, Delta := 1.0E-4, Message := 'integration resumes');
AssertEquals_WORD(Expected := 0, Actual := fbPid.stSts.stCommon.wWarning, Message := 'warning cleared');
coUnit.TEST_FINISHED();

(* ---- FirstCallReportsDevTypeAndAlarmCount.method.decl.st ---- *)
// Первый вызов: тип устройства Pid в stSts.stCommon.eDevType, один слот тревог (PID_ALARM_COUNT),
// режим из stRetain (Manual по умолчанию), Local не поддерживается (RequestMode(Local) = FALSE).
METHOD PRIVATE FirstCallReportsDevTypeAndAlarmCount
VAR
    fbTime   : FB_FakeTime;       // подменное время, старт 1 ч
    fbPid    : FB_PID;            // ФБ под тестом
    stCmd    : ST_PidCmd;         // команды
    stRetain : ST_DeviceRetain;   // режим: Manual
    stCfg    : ST_PidCfg;         // конфигурация по умолчанию
END_VAR

(* ---- FopdtClosedLoopMatchesPythonReference.method.decl.st ---- *)
// Замкнутый контур с моделью FOPDT (K = 2, T = 20 с, L = 4 с, шаг 0,1 с; параметры вымышленные):
// ПИД Kp = 1, Ti = 20 с, Td = 1 с, старт в Auto при y = 0, ступень задания 0 -> 40. Выход ПИД и PV
// в моменты 10, 30, 60, 120 с совпадают с эталоном до 1·10^-3; перерегулирование и время
// установления (полоса ±2 %) — тоже.
METHOD PRIVATE FopdtClosedLoopMatchesPythonReference
VAR
    fbTime    : FB_FakeTime;       // подменное время, старт 1 ч
    fbPid     : FB_PID;            // ФБ под тестом
    fbPlant   : FB_FopdtModel;     // модель объекта
    stCmd     : ST_PidCmd;         // команды
    stRetain  : ST_DeviceRetain;   // режим: Auto из Retain
    stCfg     : ST_PidCfg;         // конфигурация теста
    iStep     : INT;               // шаг модели (0,1 с)
    rPeak     : REAL;              // максимум PV
    rSettle_s : REAL;              // время установления, с
    rOut10    : REAL;              // выход и PV в 10, 30, 60 и 120 с
    rPv10     : REAL;
    rOut30    : REAL;
    rPv30     : REAL;
    rOut60    : REAL;
    rPv60     : REAL;
    rOut120   : REAL;
    rPv120    : REAL;
END_VAR

(* ---- FopdtClosedLoopMatchesPythonReference.method.impl.st ---- *)
coUnit.TEST('Pid_Fopdt_ClosedLoop_MatchesPythonReference');
// источник: tools/reference/pid.py, сценарий fopdt_step
stCfg.rKp := 1.0;
stCfg.rTi_s := 20.0;
stCfg.rTd_s := 1.0;
stRetain.eRemoteMode := E_DeviceMode.Auto;
stCmd.rSp_eu := 0.0;
fbPid.rPv_eu := fbPlant.rY;
fbPid.xPvValid := TRUE;
fbPid(itfTime := fbTime, stCmd := stCmd, stRetain := stRetain, stCfg := stCfg);       // t0: Auto, y = 0
stCmd.rSp_eu := 40.0;                                                                  // ступень задания
FOR iStep := 1 TO 1200 DO                                                              // 120 с
    fbTime.Advance(tStep := T#100MS);
    fbPid.rPv_eu := fbPlant.rY;
    fbPid(itfTime := fbTime, stCmd := stCmd, stRetain := stRetain, stCfg := stCfg);
    fbPlant.rU_pct := fbPid.rOut_pct;
    fbPlant.Step();
    rPeak := MAX(rPeak, fbPlant.rY);
    IF ABS(fbPlant.rY - 40.0) > 0.8 THEN                                               // вне полосы ±2 %
        rSettle_s := INT_TO_REAL(iStep + 1) * 0.1;
    END_IF
    IF iStep = 100 THEN
        rOut10 := fbPid.rOut_pct;
        rPv10 := fbPlant.rY;
    ELSIF iStep = 300 THEN
        rOut30 := fbPid.rOut_pct;
        rPv30 := fbPlant.rY;
    ELSIF iStep = 600 THEN
        rOut60 := fbPid.rOut_pct;
        rPv60 := fbPlant.rY;
    ELSIF iStep = 1200 THEN
        rOut120 := fbPid.rOut_pct;
        rPv120 := fbPlant.rY;
    END_IF
END_FOR
// ref: fopdt_step.out_10s
AssertEquals_REAL(Expected := 31.212418, Actual := rOut10, Delta := 1.0E-3, Message := 'out at 10 s');
// ref: fopdt_step.pv_10s
AssertEquals_REAL(Expected := 22.549984, Actual := rPv10, Delta := 1.0E-3, Message := 'PV at 10 s');
// ref: fopdt_step.out_30s
AssertEquals_REAL(Expected := 20.687187, Actual := rOut30, Delta := 1.0E-3, Message := 'out at 30 s');
// ref: fopdt_step.pv_30s
AssertEquals_REAL(Expected := 40.311687, Actual := rPv30, Delta := 1.0E-3, Message := 'PV at 30 s');
// ref: fopdt_step.out_60s
AssertEquals_REAL(Expected := 19.997665, Actual := rOut60, Delta := 1.0E-3, Message := 'out at 60 s');
// ref: fopdt_step.pv_60s
AssertEquals_REAL(Expected := 40.32325, Actual := rPv60, Delta := 1.0E-3, Message := 'PV at 60 s');
// ref: fopdt_step.out_120s
AssertEquals_REAL(Expected := 19.999441, Actual := rOut120, Delta := 1.0E-3, Message := 'out at 120 s');
// ref: fopdt_step.pv_120s
AssertEquals_REAL(Expected := 40.012321, Actual := rPv120, Delta := 1.0E-3, Message := 'PV at 120 s');
// ref: fopdt_step.peak
AssertEquals_REAL(Expected := 40.668068, Actual := rPeak, Delta := 1.0E-3, Message := 'peak PV');
// ref: fopdt_step.overshoot_pct
AssertEquals_REAL(Expected := 1.67017, Actual := (rPeak - 40.0) / 40.0 * 100.0, Delta := 1.0E-2,
                  Message := 'overshoot %');
// ref: fopdt_step.settle_s
AssertEquals_REAL(Expected := 24.3, Actual := rSettle_s, Delta := 0.05, Message := 'settling time, 2 % band');
coUnit.TEST_FINISHED();

(* ---- FopdtSaturatedStepBackCalcLimitsOvershoot.method.decl.st ---- *)
// Насыщение в замкнутом контуре: тот же объект и ПИД, предел выхода 30 %, ступень задания 0 -> 40,
// 60 с. С обратным расчётом (Tt = авто) выход раньше уходит с предела и перерегулирования нет;
// без него (Tt = 1·10^6 с) интегратор накапливается, перерегулирование около 9 %.
METHOD PRIVATE FopdtSaturatedStepBackCalcLimitsOvershoot
VAR
    fbTime     : FB_FakeTime;       // подменное время, старт 1 ч
    fbPidAw    : FB_PID;            // ФБ под тестом: Tt = авто
    fbPidNoAw  : FB_PID;            // сравнение: Tt = 1e6 с
    fbPlantAw  : FB_FopdtModel;     // модели объекта
    fbPlantNo  : FB_FopdtModel;
    stCmdAw    : ST_PidCmd;         // команды
    stCmdNoAw  : ST_PidCmd;
    stRetAw    : ST_DeviceRetain;   // режим: Auto из Retain
    stRetNoAw  : ST_DeviceRetain;
    stCfgAw    : ST_PidCfg;         // конфигурация
    stCfgNoAw  : ST_PidCfg;
    iStep      : INT;               // шаг модели (0,1 с)
    rPeakAw    : REAL;              // максимум PV
    rPeakNoAw  : REAL;
    xSatAw     : BOOL;              // выход был на пределе
    xSatNoAw   : BOOL;
    rUnsatAw   : REAL;              // когда выход ушёл с предела, с
    rUnsatNoAw : REAL;
END_VAR

(* ---- FopdtSaturatedStepBackCalcLimitsOvershoot.method.impl.st ---- *)
coUnit.TEST('Pid_Fopdt_SaturatedStep_BackCalcLimitsOvershoot');
// источник: tools/reference/pid.py, сценарий fopdt_sat
stCfgAw.rKp := 1.0;
stCfgAw.rTi_s := 20.0;
stCfgAw.rTd_s := 1.0;
stCfgAw.rOutMax_pct := 30.0;
stCfgNoAw := stCfgAw;
stCfgNoAw.rTt_s := 1.0E6;
stRetAw.eRemoteMode := E_DeviceMode.Auto;
stRetNoAw.eRemoteMode := E_DeviceMode.Auto;
fbPidAw.rPv_eu := fbPlantAw.rY;
fbPidAw.xPvValid := TRUE;
fbPidNoAw.rPv_eu := fbPlantNo.rY;
fbPidNoAw.xPvValid := TRUE;
fbPidAw(itfTime := fbTime, stCmd := stCmdAw, stRetain := stRetAw, stCfg := stCfgAw);          // t0: Auto
fbPidNoAw(itfTime := fbTime, stCmd := stCmdNoAw, stRetain := stRetNoAw, stCfg := stCfgNoAw);
stCmdAw.rSp_eu := 40.0;                                                                         // ступень
stCmdNoAw.rSp_eu := 40.0;
FOR iStep := 1 TO 600 DO                                                                        // 60 с
    fbTime.Advance(tStep := T#100MS);
    fbPidAw.rPv_eu := fbPlantAw.rY;
    fbPidNoAw.rPv_eu := fbPlantNo.rY;
    fbPidAw(itfTime := fbTime, stCmd := stCmdAw, stRetain := stRetAw, stCfg := stCfgAw);
    fbPidNoAw(itfTime := fbTime, stCmd := stCmdNoAw, stRetain := stRetNoAw, stCfg := stCfgNoAw);
    fbPlantAw.rU_pct := fbPidAw.rOut_pct;
    fbPlantAw.Step();
    fbPlantNo.rU_pct := fbPidNoAw.rOut_pct;
    fbPlantNo.Step();
    rPeakAw := MAX(rPeakAw, fbPlantAw.rY);
    rPeakNoAw := MAX(rPeakNoAw, fbPlantNo.rY);
    IF fbPidAw.xSatHigh THEN
        xSatAw := TRUE;
    ELSIF xSatAw AND rUnsatAw = 0.0 THEN
        rUnsatAw := INT_TO_REAL(iStep) * 0.1;
    END_IF
    IF fbPidNoAw.xSatHigh THEN
        xSatNoAw := TRUE;
    ELSIF xSatNoAw AND rUnsatNoAw = 0.0 THEN
        rUnsatNoAw := INT_TO_REAL(iStep) * 0.1;
    END_IF
END_FOR
// ref: fopdt_sat.peak_aw
AssertEquals_REAL(Expected := 39.466667, Actual := rPeakAw, Delta := 1.0E-3, Message := 'back-calculation: peak');
// ref: fopdt_sat.peak_noaw
AssertEquals_REAL(Expected := 43.642101, Actual := rPeakNoAw, Delta := 1.0E-3, Message := 'windup: peak');
// ref: fopdt_sat.pv_60s_noaw
AssertEquals_REAL(Expected := 41.619171, Actual := fbPlantNo.rY, Delta := 1.0E-3, Message := 'windup: PV at 60 s');
// ref: fopdt_sat.unsat_aw
AssertEquals_REAL(Expected := 8.4, Actual := rUnsatAw, Delta := 0.05, Message := 'back-calculation: leaves limit');
// ref: fopdt_sat.unsat_noaw
AssertEquals_REAL(Expected := 20.8, Actual := rUnsatNoAw, Delta := 0.05, Message := 'windup: leaves limit later');
AssertTrue(Condition := rPeakAw <= 40.0, Message := 'no overshoot with back-calculation');
AssertTrue(Condition := rPeakNoAw > 42.0, Message := 'overshoot without back-calculation');
coUnit.TEST_FINISHED();

(* ---- IntegralConstantErrorRampRateKpOverTi.method.decl.st ---- *)
// ПИ-регулятор (Kp = 2, Ti = 10 с) при постоянной ошибке 4 %: выход растёт со скоростью
// Kp·e/Ti = 0,8 %/с, интегратор — на Kp·dt/Ti·e за шаг.
METHOD PRIVATE IntegralConstantErrorRampRateKpOverTi
VAR
    fbTime    : FB_FakeTime;       // подменное время, старт 1 ч
    fbPid     : FB_PID;            // ФБ под тестом
    stCmd     : ST_PidCmd;         // команды
    stRetain  : ST_DeviceRetain;   // режим: старт в Manual
    stCfg     : ST_PidCfg;         // конфигурация теста
    iStep     : INT;               // шаг цикла
    rOutFirst : REAL;              // выход в первом шаге с ошибкой
END_VAR

(* ---- IntegralConstantErrorRampRateKpOverTi.method.impl.st ---- *)
coUnit.TEST('Pid_Integral_ConstantError_RampRateKpOverTi');
// источник: tools/reference/pid.py, сценарий integral
stCfg.rKp := 2.0;
stCfg.rTi_s := 10.0;
stCmd.rManualOut_pct := 30.0;
stCmd.rSp_eu := 50.0;
fbPid.rPv_eu := 50.0;
fbPid.xPvValid := TRUE;
fbPid(itfTime := fbTime, stCmd := stCmd, stRetain := stRetain, stCfg := stCfg);       // t0: Manual
fbTime.Advance(tStep := T#100MS);
stCmd.stCommon.xSetAuto := TRUE;
fbPid(itfTime := fbTime, stCmd := stCmd, stRetain := stRetain, stCfg := stCfg);       // Auto
fbPid.rPv_eu := 46.0;                                                                  // e = 4 %
fbTime.Advance(tStep := T#100MS);
fbPid(itfTime := fbTime, stCmd := stCmd, stRetain := stRetain, stCfg := stCfg);
rOutFirst := fbPid.rOut_pct;
FOR iStep := 1 TO 50 DO                                                                // ещё 5 с
    fbTime.Advance(tStep := T#100MS);
    fbPid(itfTime := fbTime, stCmd := stCmd, stRetain := stRetain, stCfg := stCfg);
END_FOR
// ref: integral.out_first
AssertEquals_REAL(Expected := 38.0, Actual := rOutFirst, Delta := 1.0E-4, Message := 'first step: P + I = 8 + 30');
// ref: integral.out_after_5s
AssertEquals_REAL(Expected := 42.0, Actual := fbPid.rOut_pct, Delta := 1.0E-4, Message := 'output after 5 s');
// ref: integral.rate_pctps
AssertEquals_REAL(Expected := 0.8, Actual := (fbPid.rOut_pct - rOutFirst) / 5.0, Delta := 1.0E-4,
                  Message := 'ramp rate Kp * e / Ti = 0.8 %/s');
// ref: integral.i_after_5s
AssertEquals_REAL(Expected := 34.08, Actual := fbPid.stSts.rI_pct, Delta := 1.0E-4, Message := 'I after 51 updates');
coUnit.TEST_FINISHED();

(* ---- InvalidCfgAtRuntimeKeepsLastValidCfg.method.decl.st ---- *)
// Cfg испорчена в работе (rKp := -1): CheckFunction, бит PID_CFG_KP, режим Auto сохраняется,
// регулирование идёт по последней корректной копии (Kp = 2).
METHOD PRIVATE InvalidCfgAtRuntimeKeepsLastValidCfg
VAR
    fbTime   : FB_FakeTime;       // подменное время, старт 1 ч
    fbPid    : FB_PID;            // ФБ под тестом
    stCmd    : ST_PidCmd;         // команды
    stRetain : ST_DeviceRetain;   // режим: старт в Manual
    stCfg    : ST_PidCfg;         // конфигурация теста
END_VAR

(* ---- InvalidCfgStartupManualOutput.method.decl.st ---- *)
// Корректной Cfg ещё не было (rKp = 0): расчёта нет, выход = LIMIT(0, rManualOut_pct, 100),
// CheckFunction, бит PID_CFG_KP, Available = FALSE; запрос Auto — RejectedCfg; слежения в Cmd
// нет (значение оператора не переписывается).
METHOD PRIVATE InvalidCfgStartupManualOutput
VAR
    fbTime   : FB_FakeTime;       // подменное время, старт 1 ч
    fbPid    : FB_PID;            // ФБ под тестом
    stCmd    : ST_PidCmd;         // команды
    stRetain : ST_DeviceRetain;   // режим: старт в Manual
    stCfg    : ST_PidCfg;         // неверная конфигурация
END_VAR

(* ---- ManualOutputClampedToLimits.method.decl.st ---- *)
// Manual: выход оператора ограничивается rOutMin_pct…rOutMax_pct (таблица 17.5), флаги насыщения
// выставляются и на самих пределах; значение оператора в Cmd ФБ не переписывает.
METHOD PRIVATE ManualOutputClampedToLimits
VAR
    fbTime   : FB_FakeTime;       // подменное время, старт 1 ч
    fbPid    : FB_PID;            // ФБ под тестом
    stCmd    : ST_PidCmd;         // команды
    stRetain : ST_DeviceRetain;   // режим
    stCfg    : ST_PidCfg;         // конфигурация теста
    rOutHi   : REAL;              // выход при 95 %
    xSatHi   : BOOL;              // xSatHigh при 95 %
    rOutLo   : REAL;              // выход при 5 %
    xSatLo   : BOOL;              // xSatLow при 5 %
END_VAR

(* ---- ManualToAutoBumpless.method.decl.st ---- *)
// Безударный переход Manual -> Auto (Kp = 2, Ti = 10 с, Td = 1 с): ошибка 3 % есть уже в
// Manual, интегратор предустановлен I = u - P - D = 35 - 6 - 0; в момент перехода выход равен
// ручному 35 %, дальше меняется только интегратором; Cmd следит за выходом в Auto.
METHOD PRIVATE ManualToAutoBumpless
VAR
    fbTime   : FB_FakeTime;       // подменное время, старт 1 ч
    fbPid    : FB_PID;            // ФБ под тестом
    stCmd    : ST_PidCmd;         // команды
    stRetain : ST_DeviceRetain;   // режим: старт в Manual
    stCfg    : ST_PidCfg;         // конфигурация теста
    iStep    : INT;               // шаг цикла
    rIManual : REAL;              // интегратор в Manual
    rOutSw   : REAL;              // выход в вызове перехода
END_VAR

(* ---- ManualToAutoBumpless.method.impl.st ---- *)
coUnit.TEST('Pid_ManualToAuto_Bumpless');
// источник: tools/reference/pid.py, сценарий manual_to_auto
stCfg.rKp := 2.0;
stCfg.rTi_s := 10.0;
stCfg.rTd_s := 1.0;
stCmd.rManualOut_pct := 35.0;
stCmd.rSp_eu := 50.0;
fbPid.rPv_eu := 47.0;                                                                  // e = 3 %
fbPid.xPvValid := TRUE;
fbPid(itfTime := fbTime, stCmd := stCmd, stRetain := stRetain, stCfg := stCfg);       // t0: Manual
FOR iStep := 1 TO 10 DO                                                                // 1 с в Manual
    fbTime.Advance(tStep := T#100MS);
    fbPid(itfTime := fbTime, stCmd := stCmd, stRetain := stRetain, stCfg := stCfg);
END_FOR
rIManual := fbPid.stSts.rI_pct;
fbTime.Advance(tStep := T#100MS);
stCmd.stCommon.xSetAuto := TRUE;
fbPid(itfTime := fbTime, stCmd := stCmd, stRetain := stRetain, stCfg := stCfg);       // Manual -> Auto
rOutSw := fbPid.rOut_pct;
FOR iStep := 1 TO 10 DO                                                                // 1 с в Auto
    fbTime.Advance(tStep := T#100MS);
    fbPid(itfTime := fbTime, stCmd := stCmd, stRetain := stRetain, stCfg := stCfg);
END_FOR
// ref: manual_to_auto.i_manual
AssertEquals_REAL(Expected := 29.0, Actual := rIManual, Delta := 1.0E-4, Message := 'I preset = u - P - D in Manual');
// ref: manual_to_auto.out_switch
AssertEquals_REAL(Expected := 35.0, Actual := rOutSw, Delta := 1.0E-4, Message := 'no bump at Manual -> Auto');
// ref: manual_to_auto.out_1s
AssertEquals_REAL(Expected := 35.599998, Actual := fbPid.rOut_pct, Delta := 1.0E-4, Message := 'then integral action');
// ref: manual_to_auto.cmd_out_1s
AssertEquals_REAL(Expected := 35.599998, Actual := stCmd.rManualOut_pct, Delta := 1.0E-4,
                  Message := 'Cmd tracks output');
AssertTrue(Condition := fbPid.Mode = E_DeviceMode.Auto, Message := 'Auto');
coUnit.TEST_FINISHED();

(* ---- OpenLoopStepMatchesPythonReference.method.decl.st ---- *)
// Модель FOPDT без регулятора: ступень входа 10 % с t = 0; первые 40 шагов (L = 4 с) выход 0,
// на 41-м шаге 0,1 = dt/T·K·u, через 24 с — по эталону (около 20·(1 - e^-1)).
METHOD PRIVATE OpenLoopStepMatchesPythonReference
VAR
    fbPlant : FB_FopdtModel;   // модель объекта (K = 2, T = 20 с по умолчанию)
    iStep   : INT;             // шаг модели (0,1 с)
    rY40    : REAL;            // выход после 40 и 41 шага
    rY41    : REAL;
END_VAR

(* ---- OpenLoopStepMatchesPythonReference.method.impl.st ---- *)
coUnit.TEST('FopdtModel_OpenLoopStep_MatchesPythonReference');
// источник: tools/reference/pid.py, сценарий fopdt_open
fbPlant.rU_pct := 10.0;
FOR iStep := 1 TO 240 DO
    fbPlant.Step();
    IF iStep = 40 THEN
        rY40 := fbPlant.rY;
    ELSIF iStep = 41 THEN
        rY41 := fbPlant.rY;
    END_IF
END_FOR
// ref: fopdt_open.y_40
AssertEquals_REAL(Expected := 0.0, Actual := rY40, Delta := 1.0E-6, Message := 'dead time 4 s: no response yet');
// ref: fopdt_open.y_41
AssertEquals_REAL(Expected := 0.1, Actual := rY41, Delta := 1.0E-6, Message := 'first response dt / T * K * u');
// ref: fopdt_open.y_240
AssertEquals_REAL(Expected := 12.660844, Actual := fbPlant.rY, Delta := 1.0E-4, Message := 'response after 24 s');
coUnit.TEST_FINISHED();

(* ---- OutOfServiceHoldsOutput.method.decl.st ---- *)
// OutOfService: выход удерживается при любой PV, расчёта нет, Cmd следит за выходом, CheckFunction;
// выход в Auto — шаг инициализации без бита DT_GAP, регулирование продолжается с удержанного
// выхода без рывка.
METHOD PRIVATE OutOfServiceHoldsOutput
VAR
    fbTime   : FB_FakeTime;       // подменное время, старт 1 ч
    fbPid    : FB_PID;            // ФБ под тестом
    stCmd    : ST_PidCmd;         // команды
    stRetain : ST_DeviceRetain;   // режим: старт в Manual
    stCfg    : ST_PidCfg;         // конфигурация теста
    iStep    : INT;               // шаг цикла
    rOutOos  : REAL;              // выход в вызове входа в OOS
    eResOos  : E_CmdResult;       // результат xSetOos
    rOutExit : REAL;              // выход в вызове выхода из OOS
    wWrnExit : WORD;              // wWarning в вызове выхода
END_VAR

(* ---- OutOfServiceHoldsOutput.method.impl.st ---- *)
coUnit.TEST('Pid_OutOfService_HoldsOutput');
// источник: tools/reference/pid.py, сценарий oos
stCfg.rKp := 2.0;
stCfg.rTi_s := 10.0;
stCmd.rManualOut_pct := 30.0;
stCmd.rSp_eu := 50.0;
fbPid.rPv_eu := 50.0;
fbPid.xPvValid := TRUE;
fbPid(itfTime := fbTime, stCmd := stCmd, stRetain := stRetain, stCfg := stCfg);       // t0: Manual
fbTime.Advance(tStep := T#100MS);
stCmd.stCommon.xSetAuto := TRUE;
fbPid(itfTime := fbTime, stCmd := stCmd, stRetain := stRetain, stCfg := stCfg);       // Auto
fbPid.rPv_eu := 46.0;                                                                  // e = 4 %
FOR iStep := 1 TO 10 DO
    fbTime.Advance(tStep := T#100MS);
    fbPid(itfTime := fbTime, stCmd := stCmd, stRetain := stRetain, stCfg := stCfg);
END_FOR
fbTime.Advance(tStep := T#100MS);
stCmd.stCommon.xSetOos := TRUE;
fbPid(itfTime := fbTime, stCmd := stCmd, stRetain := stRetain, stCfg := stCfg);       // в OutOfService
rOutOos := fbPid.rOut_pct;
eResOos := fbPid.stSts.stCommon.eCmdResult;
fbPid.rPv_eu := 30.0;                                                                  // PV меняется
FOR iStep := 1 TO 30 DO
    fbTime.Advance(tStep := T#100MS);
    fbPid(itfTime := fbTime, stCmd := stCmd, stRetain := stRetain, stCfg := stCfg);
END_FOR
// ref: oos.out_oos
AssertEquals_REAL(Expected := 38.72, Actual := rOutOos, Delta := 1.0E-4, Message := 'OOS entry keeps output');
AssertTrue(Condition := eResOos = E_CmdResult.Accepted, Message := 'xSetOos accepted');
// ref: oos.out_oos_3s
AssertEquals_REAL(Expected := 38.72, Actual := fbPid.rOut_pct, Delta := 1.0E-4, Message := 'held in OOS');
AssertEquals_REAL(Expected := 38.72, Actual := stCmd.rManualOut_pct, Delta := 1.0E-4, Message := 'Cmd tracks output');
AssertTrue(Condition := fbPid.Status = E_Ne107Status.CheckFunction, Message := 'CheckFunction in OOS');
AssertTrue(Condition := stRetain.xOutOfService, Message := 'OOS in retain');
fbTime.Advance(tStep := T#100MS);
stCmd.stCommon.xSetAuto := TRUE;
fbPid(itfTime := fbTime, stCmd := stCmd, stRetain := stRetain, stCfg := stCfg);       // выход из OOS
rOutExit := fbPid.rOut_pct;
wWrnExit := fbPid.stSts.stCommon.wWarning;
FOR iStep := 1 TO 2 DO
    fbTime.Advance(tStep := T#100MS);
    fbPid(itfTime := fbTime, stCmd := stCmd, stRetain := stRetain, stCfg := stCfg);
END_FOR
// ref: oos.out_exit
AssertEquals_REAL(Expected := 38.72, Actual := rOutExit, Delta := 1.0E-4, Message := 'no bump on OOS exit');
AssertEquals_WORD(Expected := 0, Actual := wWrnExit, Message := 'OOS exit is not a time gap');
// ref: oos.out_exit_2
AssertEquals_REAL(Expected := 39.12, Actual := fbPid.rOut_pct, Delta := 1.0E-4, Message := 'control resumes, e = 20 %');
coUnit.TEST_FINISHED();

(* ---- OutputLimitsClampAndFlags.method.decl.st ---- *)
// Пределы выхода 10…90 % (Kp = 2, без I): большая положительная ошибка — выход 90 % и xSatHigh
// (бит SAT_HIGH), большая отрицательная — 10 % и xSatLow (бит SAT_LOW).
METHOD PRIVATE OutputLimitsClampAndFlags
VAR
    fbTime   : FB_FakeTime;       // подменное время, старт 1 ч
    fbPid    : FB_PID;            // ФБ под тестом
    stCmd    : ST_PidCmd;         // команды
    stRetain : ST_DeviceRetain;   // режим: старт в Manual
    stCfg    : ST_PidCfg;         // конфигурация теста
END_VAR

(* ---- OutputRateLimitIntegratorBacksOff.method.decl.st ---- *)
// Ограничение скорости выхода 5 %/с (Kp = 2, Ti = 10 с): после ступени задания на 10 % выход
// растёт ровно на 0,5 % за шаг 100 мс (бит OUT_RATE_LIMITED), а обратный расчёт по разности
// u - v сдерживает интегратор (без него было бы 40 + 2·10·2/10 = 44 % за 2 с).
METHOD PRIVATE OutputRateLimitIntegratorBacksOff
VAR
    fbTime   : FB_FakeTime;       // подменное время, старт 1 ч
    fbPid    : FB_PID;            // ФБ под тестом
    stCmd    : ST_PidCmd;         // команды
    stRetain : ST_DeviceRetain;   // режим: старт в Manual
    stCfg    : ST_PidCfg;         // конфигурация теста
    iStep    : INT;               // шаг цикла
END_VAR

(* ---- OutputRateLimitIntegratorBacksOff.method.impl.st ---- *)
coUnit.TEST('Pid_OutputRateLimit_IntegratorBacksOff');
// источник: tools/reference/pid.py, сценарий rate_limit
stCfg.rKp := 2.0;
stCfg.rTi_s := 10.0;
stCfg.rOutRate_pctps := 5.0;
stCmd.rManualOut_pct := 40.0;
stCmd.rSp_eu := 50.0;
fbPid.rPv_eu := 50.0;
fbPid.xPvValid := TRUE;
fbPid(itfTime := fbTime, stCmd := stCmd, stRetain := stRetain, stCfg := stCfg);       // t0: Manual
fbTime.Advance(tStep := T#100MS);
stCmd.stCommon.xSetAuto := TRUE;
fbPid(itfTime := fbTime, stCmd := stCmd, stRetain := stRetain, stCfg := stCfg);       // Auto
stCmd.rSp_eu := 60.0;                                                                  // P: 0 -> 20 %
FOR iStep := 1 TO 20 DO                                                                // 2 с
    fbTime.Advance(tStep := T#100MS);
    fbPid(itfTime := fbTime, stCmd := stCmd, stRetain := stRetain, stCfg := stCfg);
END_FOR
// ref: rate_limit.out_2s
AssertEquals_REAL(Expected := 50.0, Actual := fbPid.rOut_pct, Delta := 1.0E-4, Message := 'out = 40 + 5 %/s * 2 s');
// ref: rate_limit.i_2s
AssertEquals_REAL(Expected := 40.986393, Actual := fbPid.stSts.rI_pct, Delta := 1.0E-3, Message := 'I backs off');
AssertTrue(Condition := fbPid.stSts.rI_pct < 44.0, Message := 'I below plain integration 44 %');
AssertEquals_WORD(Expected := GVL_Const.PID_STS_OUT_RATE_LIMITED,
                  Actual := fbPid.stSts.stCommon.wStatus AND GVL_Const.PID_STS_OUT_RATE_LIMITED,
                  Message := 'status bit OUT_RATE_LIMITED');
coUnit.TEST_FINISHED();

(* ---- POnlyErrorStepOutputEqualsKpTimesError.method.decl.st ---- *)
// П-регулятор (Kp = 2, без I и D): после безударного перехода в Auto со смещением 40 % выход
// отличается от смещения ровно на Kp·e при ошибке +5 % и -3 %.
METHOD PRIVATE POnlyErrorStepOutputEqualsKpTimesError
VAR
    fbTime   : FB_FakeTime;       // подменное время, старт 1 ч
    fbPid    : FB_PID;            // ФБ под тестом
    stCmd    : ST_PidCmd;         // команды
    stRetain : ST_DeviceRetain;   // режим: старт в Manual
    stCfg    : ST_PidCfg;         // конфигурация теста
END_VAR

(* ---- PvFailHoldOutputBumplessResume.method.decl.st ---- *)
// Отказ PV в Auto, реакция Hold (Kp = 2, Ti = 10 с): выход удерживается, интегратор заморожен,
// Failure, бит PID_FLT_PV_INVALID, бит PV_FAIL, тревога PvInvalid активна. PV вернулась с другой
// ошибкой (6 % вместо 4 %): шаг инициализации, выход продолжается с удержанного без рывка.
METHOD PRIVATE PvFailHoldOutputBumplessResume
VAR
    fbTime   : FB_FakeTime;       // подменное время, старт 1 ч
    fbPid    : FB_PID;            // ФБ под тестом
    stCmd    : ST_PidCmd;         // команды
    stRetain : ST_DeviceRetain;   // режим: старт в Manual
    stCfg    : ST_PidCfg;         // конфигурация теста
    iStep    : INT;               // шаг цикла
    rBefore  : REAL;              // выход до отказа
    rFail    : REAL;              // выход через 2 с отказа
    eStFail  : E_Ne107Status;     // статус при отказе
    wFltFail : WORD;              // wFault при отказе
    wStsFail : WORD;              // wStatus при отказе
    wAlmFail : WORD;              // wAlmActive при отказе
    rResume  : REAL;              // выход в вызове возврата PV
END_VAR

(* ---- PvFailHoldOutputBumplessResume.method.impl.st ---- *)
coUnit.TEST('Pid_PvFail_HoldOutput_BumplessResume');
// источник: tools/reference/pid.py, сценарий pv_fail_hold
stCfg.rKp := 2.0;
stCfg.rTi_s := 10.0;
stCmd.rManualOut_pct := 30.0;
stCmd.rSp_eu := 50.0;
fbPid.rPv_eu := 50.0;
fbPid.xPvValid := TRUE;
fbPid(itfTime := fbTime, stCmd := stCmd, stRetain := stRetain, stCfg := stCfg);       // t0: Manual
fbTime.Advance(tStep := T#100MS);
stCmd.stCommon.xSetAuto := TRUE;
fbPid(itfTime := fbTime, stCmd := stCmd, stRetain := stRetain, stCfg := stCfg);       // Auto
fbPid.rPv_eu := 46.0;                                                                  // e = 4 %
FOR iStep := 1 TO 10 DO
    fbTime.Advance(tStep := T#100MS);
    fbPid(itfTime := fbTime, stCmd := stCmd, stRetain := stRetain, stCfg := stCfg);
END_FOR
rBefore := fbPid.rOut_pct;
fbPid.xPvValid := FALSE;                                                               // отказ PV
FOR iStep := 1 TO 20 DO
    fbTime.Advance(tStep := T#100MS);
    fbPid(itfTime := fbTime, stCmd := stCmd, stRetain := stRetain, stCfg := stCfg);
END_FOR
rFail := fbPid.rOut_pct;
eStFail := fbPid.Status;
wFltFail := fbPid.stSts.stCommon.wFault;
wStsFail := fbPid.stSts.stCommon.wStatus;
wAlmFail := fbPid.stSts.stCommon.wAlmActive;
fbPid.xPvValid := TRUE;                                                                // PV вернулась
fbPid.rPv_eu := 44.0;                                                                  // e = 6 %
fbTime.Advance(tStep := T#100MS);
fbPid(itfTime := fbTime, stCmd := stCmd, stRetain := stRetain, stCfg := stCfg);
rResume := fbPid.rOut_pct;
FOR iStep := 1 TO 2 DO
    fbTime.Advance(tStep := T#100MS);
    fbPid(itfTime := fbTime, stCmd := stCmd, stRetain := stRetain, stCfg := stCfg);
END_FOR
// ref: pv_fail_hold.out_before
AssertEquals_REAL(Expected := 38.72, Actual := rBefore, Delta := 1.0E-4, Message := 'output before PV failure');
// ref: pv_fail_hold.out_fail
AssertEquals_REAL(Expected := 38.72, Actual := rFail, Delta := 1.0E-4, Message := 'Hold: output held');
AssertTrue(Condition := eStFail = E_Ne107Status.Failure, Message := 'Failure while PV invalid in Auto');
AssertEquals_WORD(Expected := GVL_Const.PID_FLT_PV_INVALID, Actual := wFltFail, Message := 'wFault PV_INVALID');
AssertEquals_WORD(Expected := GVL_Const.PID_STS_PV_FAIL, Actual := wStsFail AND GVL_Const.PID_STS_PV_FAIL,
                  Message := 'status bit PV_FAIL');
AssertEquals_WORD(Expected := 16#0001, Actual := wAlmFail, Message := 'alarm PvInvalid active');
// ref: pv_fail_hold.out_resume
AssertEquals_REAL(Expected := 38.72, Actual := rResume, Delta := 1.0E-4, Message := 'resume without bump');
// ref: pv_fail_hold.out_resume_2
AssertEquals_REAL(Expected := 38.84, Actual := fbPid.rOut_pct, Delta := 1.0E-4,
                  Message := 'then integral with e = 6 %');
AssertTrue(Condition := fbPid.Status = E_Ne107Status.Good, Message := 'Good after PV recovery');
coUnit.TEST_FINISHED();

(* ---- PvFailSafeOutDrivesSafeOutput.method.decl.st ---- *)
// Отказ PV в Auto, реакция SafeOut (rSafeOut_pct = 15 %): выход 15 % без рампы; после возврата PV
// регулирование продолжается с 15 % без рывка (шаг инициализации).
METHOD PRIVATE PvFailSafeOutDrivesSafeOutput
VAR
    fbTime   : FB_FakeTime;       // подменное время, старт 1 ч
    fbPid    : FB_PID;            // ФБ под тестом
    stCmd    : ST_PidCmd;         // команды
    stRetain : ST_DeviceRetain;   // режим: старт в Manual
    stCfg    : ST_PidCfg;         // конфигурация теста
    iStep    : INT;               // шаг цикла
    rFail    : REAL;              // выход при отказе
    rResume  : REAL;              // выход в вызове возврата PV
END_VAR

(* ---- PvFailSafeOutDrivesSafeOutput.method.impl.st ---- *)
coUnit.TEST('Pid_PvFail_SafeOut_DrivesSafeOutput');
// источник: tools/reference/pid.py, сценарий safe_out
stCfg.rKp := 2.0;
stCfg.rTi_s := 10.0;
stCfg.ePvFailAction := E_PidPvFailAction.SafeOut;
stCfg.rSafeOut_pct := 15.0;
stCmd.rManualOut_pct := 30.0;
stCmd.rSp_eu := 50.0;
fbPid.rPv_eu := 50.0;
fbPid.xPvValid := TRUE;
fbPid(itfTime := fbTime, stCmd := stCmd, stRetain := stRetain, stCfg := stCfg);       // t0: Manual
fbTime.Advance(tStep := T#100MS);
stCmd.stCommon.xSetAuto := TRUE;
fbPid(itfTime := fbTime, stCmd := stCmd, stRetain := stRetain, stCfg := stCfg);       // Auto
fbPid.rPv_eu := 46.0;                                                                  // e = 4 %
FOR iStep := 1 TO 10 DO
    fbTime.Advance(tStep := T#100MS);
    fbPid(itfTime := fbTime, stCmd := stCmd, stRetain := stRetain, stCfg := stCfg);
END_FOR
fbPid.xPvValid := FALSE;                                                               // отказ PV
FOR iStep := 1 TO 5 DO
    fbTime.Advance(tStep := T#100MS);
    fbPid(itfTime := fbTime, stCmd := stCmd, stRetain := stRetain, stCfg := stCfg);
END_FOR
rFail := fbPid.rOut_pct;
fbPid.xPvValid := TRUE;                                                                // PV вернулась
fbTime.Advance(tStep := T#100MS);
fbPid(itfTime := fbTime, stCmd := stCmd, stRetain := stRetain, stCfg := stCfg);
rResume := fbPid.rOut_pct;
FOR iStep := 1 TO 2 DO
    fbTime.Advance(tStep := T#100MS);
    fbPid(itfTime := fbTime, stCmd := stCmd, stRetain := stRetain, stCfg := stCfg);
END_FOR
// ref: safe_out.out_fail
AssertEquals_REAL(Expected := 15.0, Actual := rFail, Delta := 1.0E-4, Message := 'SafeOut: rSafeOut_pct');
// ref: safe_out.out_resume
AssertEquals_REAL(Expected := 15.0, Actual := rResume, Delta := 1.0E-4, Message := 'resume from safe output');
// ref: safe_out.out_resume_2
AssertEquals_REAL(Expected := 15.08, Actual := fbPid.rOut_pct, Delta := 1.0E-4, Message := 'then integral action');
AssertTrue(Condition := fbPid.Mode = E_DeviceMode.Auto, Message := 'stays Auto');
coUnit.TEST_FINISHED();

(* ---- PvFailShedToManual.method.decl.st ---- *)
// Отказ PV в Auto, реакция ShedToManual: ФБ переходит в Manual (и в stRetain) с текущим выходом,
// stCmd.rManualOut_pct уже равен выходу; в Manual отказ PV — не Failure.
METHOD PRIVATE PvFailShedToManual
VAR
    fbTime   : FB_FakeTime;       // подменное время, старт 1 ч
    fbPid    : FB_PID;            // ФБ под тестом
    stCmd    : ST_PidCmd;         // команды
    stRetain : ST_DeviceRetain;   // режим: старт в Manual
    stCfg    : ST_PidCfg;         // конфигурация теста
    iStep    : INT;               // шаг цикла
END_VAR

(* ---- PvFailShedToManual.method.impl.st ---- *)
coUnit.TEST('Pid_PvFail_ShedToManual');
// источник: tools/reference/pid.py, сценарий pv_fail_hold (та же последовательность до отказа)
stCfg.rKp := 2.0;
stCfg.rTi_s := 10.0;
stCfg.ePvFailAction := E_PidPvFailAction.ShedToManual;
stCmd.rManualOut_pct := 30.0;
stCmd.rSp_eu := 50.0;
fbPid.rPv_eu := 50.0;
fbPid.xPvValid := TRUE;
fbPid(itfTime := fbTime, stCmd := stCmd, stRetain := stRetain, stCfg := stCfg);       // t0: Manual
fbTime.Advance(tStep := T#100MS);
stCmd.stCommon.xSetAuto := TRUE;
fbPid(itfTime := fbTime, stCmd := stCmd, stRetain := stRetain, stCfg := stCfg);       // Auto
fbPid.rPv_eu := 46.0;                                                                  // e = 4 %
FOR iStep := 1 TO 10 DO
    fbTime.Advance(tStep := T#100MS);
    fbPid(itfTime := fbTime, stCmd := stCmd, stRetain := stRetain, stCfg := stCfg);
END_FOR
fbPid.xPvValid := FALSE;                                                               // отказ PV
fbTime.Advance(tStep := T#100MS);
fbPid(itfTime := fbTime, stCmd := stCmd, stRetain := stRetain, stCfg := stCfg);
AssertTrue(Condition := fbPid.Mode = E_DeviceMode.Manual, Message := 'shed to Manual');
AssertTrue(Condition := stRetain.eRemoteMode = E_DeviceMode.Manual, Message := 'Manual remembered in retain');
// ref: pv_fail_hold.out_before
AssertEquals_REAL(Expected := 38.72, Actual := fbPid.rOut_pct, Delta := 1.0E-4, Message := 'keeps current output');
AssertEquals_REAL(Expected := 38.72, Actual := stCmd.rManualOut_pct, Delta := 1.0E-4,
                  Message := 'Cmd holds the output');
AssertTrue(Condition := fbPid.Status = E_Ne107Status.Good, Message := 'no Failure in Manual');
AssertEquals_WORD(Expected := 0, Actual := fbPid.stSts.stCommon.wFault, Message := 'wFault 0 in Manual');
coUnit.TEST_FINISHED();

(* ---- PvFailShedToManualAlarmStaysActive.method.decl.st ---- *)
// Отказ PV в Auto с реакцией ShedToManual: ФБ сам уходит в Manual, и тревога PvInvalid всё равно
// появляется (ActiveUnack) и держится, пока PV негодна: оператор должен узнать, что контур
// переведён на ручное управление. Возврат PV снимает условие (RtnUnack), квитирование — Normal.
// Выход из OutOfService в Manual при негодной PV тревоги не даёт: Manual выбрал оператор.
METHOD PRIVATE PvFailShedToManualAlarmStaysActive
VAR
    fbTime   : FB_FakeTime;       // подменное время, старт 1 ч
    fbPid    : FB_PID;            // ФБ под тестом
    stCmd    : ST_PidCmd;         // команды
    stRetain : ST_DeviceRetain;   // режим: старт в Manual
    stCfg    : ST_PidCfg;         // конфигурация теста
    itfAlm   : I_Alarm;           // тревога PvInvalid
    iStep    : INT;               // шаг цикла
    eModeSh  : E_DeviceMode;      // режим в вызове отказа PV
    eStShed  : E_AlarmState;      // тревога в вызове отказа PV
    eStHeld  : E_AlarmState;      // через 5 с в Manual при негодной PV
    wActHeld : WORD;              // wAlmActive через 5 с
    wUnaHeld : WORD;              // wAlmUnack через 5 с
    eStRtn   : E_AlarmState;      // после возврата PV
    eStAck   : E_AlarmState;      // после квитирования
    eStOper  : E_AlarmState;      // OutOfService -> Manual оператором при негодной PV
END_VAR

(* ---- PvFailShedToManualAlarmStaysActive.method.impl.st ---- *)
coUnit.TEST('Pid_PvFail_ShedToManual_AlarmStaysActive');
stCfg.ePvFailAction := E_PidPvFailAction.ShedToManual;
stCfg.udiAlarmIdBase := 70;
stCmd.rManualOut_pct := 30.0;
stCmd.rSp_eu := 50.0;
fbPid.rPv_eu := 50.0;
fbPid.xPvValid := TRUE;
fbPid(itfTime := fbTime, stCmd := stCmd, stRetain := stRetain, stCfg := stCfg);       // t0: Manual
itfAlm := fbPid.GetAlarm(uiIndex := TO_UINT(E_PidAlarm.PvInvalid));
fbTime.Advance(tStep := T#100MS);
stCmd.stCommon.xSetAuto := TRUE;
fbPid(itfTime := fbTime, stCmd := stCmd, stRetain := stRetain, stCfg := stCfg);       // Auto
fbPid.xPvValid := FALSE;                                                               // отказ PV
fbTime.Advance(tStep := T#100MS);
fbPid(itfTime := fbTime, stCmd := stCmd, stRetain := stRetain, stCfg := stCfg);       // сброс в Manual
eModeSh := fbPid.Mode;
eStShed := itfAlm.State;
FOR iStep := 1 TO 50 DO                                                                // 5 с, PV негодна
    fbTime.Advance(tStep := T#100MS);
    fbPid(itfTime := fbTime, stCmd := stCmd, stRetain := stRetain, stCfg := stCfg);
END_FOR
eStHeld := itfAlm.State;
wActHeld := fbPid.stSts.stCommon.wAlmActive;
wUnaHeld := fbPid.stSts.stCommon.wAlmUnack;
fbPid.xPvValid := TRUE;                                                                // PV вернулась
fbTime.Advance(tStep := T#100MS);
fbPid(itfTime := fbTime, stCmd := stCmd, stRetain := stRetain, stCfg := stCfg);
eStRtn := itfAlm.State;
stCmd.stCommon.xAck := TRUE;
fbTime.Advance(tStep := T#100MS);
fbPid(itfTime := fbTime, stCmd := stCmd, stRetain := stRetain, stCfg := stCfg);
eStAck := itfAlm.State;
// Manual после OutOfService выбрал оператор: негодная PV тревоги не даёт
stCmd.stCommon.xSetOos := TRUE;
fbTime.Advance(tStep := T#100MS);
fbPid(itfTime := fbTime, stCmd := stCmd, stRetain := stRetain, stCfg := stCfg);
fbPid.xPvValid := FALSE;
stCmd.stCommon.xSetManual := TRUE;
fbTime.Advance(tStep := T#100MS);
fbPid(itfTime := fbTime, stCmd := stCmd, stRetain := stRetain, stCfg := stCfg);
fbTime.Advance(tStep := T#100MS);
fbPid(itfTime := fbTime, stCmd := stCmd, stRetain := stRetain, stCfg := stCfg);
eStOper := itfAlm.State;
AssertTrue(Condition := eModeSh = E_DeviceMode.Manual, Message := 'shed to Manual');
AssertTrue(Condition := eStShed = E_AlarmState.ActiveUnack, Message := 'alarm ActiveUnack in the shed call');
AssertTrue(Condition := eStHeld = E_AlarmState.ActiveUnack, Message := 'alarm stays active while PV is invalid');
AssertEquals_WORD(Expected := 16#0001, Actual := wActHeld, Message := 'wAlmActive slot 0 while PV is invalid');
AssertEquals_WORD(Expected := 16#0001, Actual := wUnaHeld, Message := 'wAlmUnack slot 0 while PV is invalid');
AssertTrue(Condition := eStRtn = E_AlarmState.RtnUnack, Message := 'RtnUnack after PV recovery');
AssertTrue(Condition := eStAck = E_AlarmState.Normal, Message := 'Normal after xAck');
AssertTrue(Condition := eStOper = E_AlarmState.Normal, Message := 'no alarm in operator-selected Manual');
coUnit.TEST_FINISHED();

(* ---- PvFailShedToManualDeferredWhileTracking.method.decl.st ---- *)
// ShedToManual при слежении не выполняется: регулятор не управляет, выход задаёт механизм. Когда
// слежение снято, а PV всё ещё негодна, — переход в Manual с текущим (отслеженным) выходом.
METHOD PRIVATE PvFailShedToManualDeferredWhileTracking
VAR
    fbTime   : FB_FakeTime;       // подменное время, старт 1 ч
    fbPid    : FB_PID;            // ФБ под тестом
    stCmd    : ST_PidCmd;         // команды
    stRetain : ST_DeviceRetain;   // режим
    stCfg    : ST_PidCfg;         // конфигурация теста
    iStep    : INT;               // шаг цикла
    eModeTrk : E_DeviceMode;      // режим через 1 с слежения
END_VAR

(* ---- PvFailShedToManualDeferredWhileTracking.method.impl.st ---- *)
coUnit.TEST('Pid_PvFail_ShedToManual_DeferredWhileTracking');
stCfg.ePvFailAction := E_PidPvFailAction.ShedToManual;
stRetain.eRemoteMode := E_DeviceMode.Auto;
stCmd.rSp_eu := 50.0;
fbPid.rPv_eu := 50.0;
fbPid.xPvValid := FALSE;
fbPid.xTrack := TRUE;
fbPid.rTrack_pct := 33.0;
fbPid(itfTime := fbTime, stCmd := stCmd, stRetain := stRetain, stCfg := stCfg);       // t0: Auto, слежение, PV негодна
FOR iStep := 1 TO 10 DO
    fbTime.Advance(tStep := T#100MS);
    fbPid(itfTime := fbTime, stCmd := stCmd, stRetain := stRetain, stCfg := stCfg);
END_FOR
eModeTrk := fbPid.Mode;
fbPid.xTrack := FALSE;                                                                 // слежение снято
fbTime.Advance(tStep := T#100MS);
fbPid(itfTime := fbTime, stCmd := stCmd, stRetain := stRetain, stCfg := stCfg);
AssertTrue(Condition := eModeTrk = E_DeviceMode.Auto, Message := 'stays Auto while tracking');
AssertTrue(Condition := fbPid.Mode = E_DeviceMode.Manual, Message := 'shed once tracking ends');
AssertTrue(Condition := stRetain.eRemoteMode = E_DeviceMode.Manual, Message := 'Manual in retain');
AssertEquals_REAL(Expected := 33.0, Actual := fbPid.rOut_pct, Delta := 0.0, Message := 'keeps tracked output');
AssertEquals_REAL(Expected := 33.0, Actual := stCmd.rManualOut_pct, Delta := 0.0, Message := 'Cmd holds the output');
coUnit.TEST_FINISHED();

(* ---- PvInvalidAlarmActiveOnlyInAuto.method.decl.st ---- *)
// Тревога слота 0 PvInvalid: в Manual негодная PV тревоги не даёт; в Auto — ActiveUnack с номером
// udiAlarmIdBase + 0, квитирование — ActiveAck, возврат PV — Normal.
METHOD PRIVATE PvInvalidAlarmActiveOnlyInAuto
VAR
    fbTime   : FB_FakeTime;       // подменное время, старт 1 ч
    fbPid    : FB_PID;            // ФБ под тестом
    stCmd    : ST_PidCmd;         // команды
    stRetain : ST_DeviceRetain;   // режим: старт в Manual
    stCfg    : ST_PidCfg;         // конфигурация теста
    itfAlm   : I_Alarm;           // тревога PvInvalid
    eStMan   : E_AlarmState;      // состояние тревоги в Manual
    eStAuto  : E_AlarmState;      // в Auto при отказе PV
    eStAck   : E_AlarmState;      // после квитирования
END_VAR

(* ---- PvNaNEventAndStsFinite.method.decl.st ---- *)
// Auto, PV = NaN при xPvValid = TRUE (мусор Modbus): тревога PvInvalid; значение её события и stSts.rPv_eu конечны —
// 0.0 (R6), выход удерживается (Hold) и конечен.
METHOD PRIVATE PvNaNEventAndStsFinite
VAR
    fbTime   : FB_FakeTime;       // подменное время, старт 1 ч
    fbPid    : FB_PID;            // ФБ под тестом
    stCmd    : ST_PidCmd;         // команды
    stRetain : ST_DeviceRetain;   // режим: Auto из Retain
    stCfg    : ST_PidCfg;         // конфигурация (умолчания)
    fbSink   : FB_TestSink;       // приёмник событий
    stEv     : ST_AlarmEvent;     // последнее событие
    uBits    : U_RealBits;        // NaN по битам
END_VAR

(* ---- PvNaNTreatedAsInvalid.method.decl.st ---- *)
// PV не конечна при xPvValid = TRUE (P-04): в Auto это отказ PV — Failure, бит PV_FAIL, wFault,
// тревога; выход удерживается (Hold), NaN в расчёт не попадает. Годная PV — продолжение без рывка.
METHOD PRIVATE PvNaNTreatedAsInvalid
VAR
    fbTime   : FB_FakeTime;       // подменное время, старт 1 ч
    fbPid    : FB_PID;            // ФБ под тестом
    stCmd    : ST_PidCmd;         // команды
    stRetain : ST_DeviceRetain;   // режим
    stCfg    : ST_PidCfg;         // конфигурация теста
    uBits    : U_RealBits;        // источник NaN
    eStNaN   : E_Ne107Status;     // статус при NaN
    wStsNaN  : WORD;              // wStatus при NaN
    wFltNaN  : WORD;              // wFault при NaN
    wAlmNaN  : WORD;              // wAlmActive при NaN
    rOutNaN  : REAL;              // выход при NaN
END_VAR

(* ---- RealDtSameResultFor10msAnd100msSteps.method.decl.st ---- *)
// Расчёт по реальному dt (Kp = 2, Ti = 10 с, e = 4 %): за 5 с при вызовах раз в 10 мс и раз в
// 100 мс интегратор одинаков (30 + 2·4·5/10 = 34 %). Выход берёт интегратор прошлого шага,
// поэтому выходы различаются ровно на приращение одного шага: 0,008 и 0,08 %.
METHOD PRIVATE RealDtSameResultFor10msAnd100msSteps
VAR
    fbTimeA  : FB_FakeTime;       // время ФБ A (шаг 10 мс)
    fbTimeB  : FB_FakeTime;       // время ФБ B (шаг 100 мс)
    fbPidA   : FB_PID;            // вызовы раз в 10 мс
    fbPidB   : FB_PID;            // вызовы раз в 100 мс
    stCmdA   : ST_PidCmd;         // команды
    stCmdB   : ST_PidCmd;
    stRetA   : ST_DeviceRetain;   // режим: старт в Manual
    stRetB   : ST_DeviceRetain;
    stCfg    : ST_PidCfg;         // общая конфигурация
    iStep    : INT;               // шаг цикла
END_VAR

(* ---- RealDtSameResultFor10msAnd100msSteps.method.impl.st ---- *)
coUnit.TEST('Pid_RealDt_SameResultFor10msAnd100msSteps');
// источник: tools/reference/pid.py, сценарий real_dt
stCfg.rKp := 2.0;
stCfg.rTi_s := 10.0;
stCmdA.rManualOut_pct := 30.0;
stCmdA.rSp_eu := 50.0;
stCmdB := stCmdA;
fbPidA.rPv_eu := 50.0;
fbPidA.xPvValid := TRUE;
fbPidB.rPv_eu := 50.0;
fbPidB.xPvValid := TRUE;
fbPidA(itfTime := fbTimeA, stCmd := stCmdA, stRetain := stRetA, stCfg := stCfg);      // t0: Manual
fbPidB(itfTime := fbTimeB, stCmd := stCmdB, stRetain := stRetB, stCfg := stCfg);
fbTimeA.Advance(tStep := T#10MS);
fbTimeB.Advance(tStep := T#100MS);
stCmdA.stCommon.xSetAuto := TRUE;
stCmdB.stCommon.xSetAuto := TRUE;
fbPidA(itfTime := fbTimeA, stCmd := stCmdA, stRetain := stRetA, stCfg := stCfg);      // Auto
fbPidB(itfTime := fbTimeB, stCmd := stCmdB, stRetain := stRetB, stCfg := stCfg);
fbPidA.rPv_eu := 46.0;                                                                 // e = 4 %
fbPidB.rPv_eu := 46.0;
FOR iStep := 1 TO 500 DO                                                               // 5 с по 10 мс
    fbTimeA.Advance(tStep := T#10MS);
    fbPidA(itfTime := fbTimeA, stCmd := stCmdA, stRetain := stRetA, stCfg := stCfg);
END_FOR
FOR iStep := 1 TO 50 DO                                                                // 5 с по 100 мс
    fbTimeB.Advance(tStep := T#100MS);
    fbPidB(itfTime := fbTimeB, stCmd := stCmdB, stRetain := stRetB, stCfg := stCfg);
END_FOR
// ref: real_dt.i_10ms
AssertEquals_REAL(Expected := 34.0, Actual := fbPidA.stSts.rI_pct, Delta := 1.0E-4,
                  Message := 'I after 5 s, 10 ms steps');
// ref: real_dt.i_100ms
AssertEquals_REAL(Expected := 34.0, Actual := fbPidB.stSts.rI_pct, Delta := 1.0E-4,
                  Message := 'I after 5 s, 100 ms steps');
AssertEquals_REAL(Expected := fbPidB.stSts.rI_pct, Actual := fbPidA.stSts.rI_pct, Delta := 1.0E-4,
                  Message := 'same integral for both cycle times');
// ref: real_dt.out_10ms
AssertEquals_REAL(Expected := 41.992001, Actual := fbPidA.rOut_pct, Delta := 1.0E-4, Message := 'out, 10 ms steps');
// ref: real_dt.out_100ms
AssertEquals_REAL(Expected := 41.919998, Actual := fbPidB.rOut_pct, Delta := 1.0E-4, Message := 'out, 100 ms steps');
coUnit.TEST_FINISHED();

(* ---- ResetAcceptedWithoutLatchedFaults.method.decl.st ---- *)
// Reset у ПИД (фиксируемых отказов нет): xReset и Reset() принимаются, каждая команда даёт +1 к
// uiCmdSeq, бит xReset сбрасывается (чек-лист устройства, пункт 2).
METHOD PRIVATE ResetAcceptedWithoutLatchedFaults
VAR
    fbTime   : FB_FakeTime;       // подменное время, старт 1 ч
    fbPid    : FB_PID;            // ФБ под тестом
    stCmd    : ST_PidCmd;         // команды
    stRetain : ST_DeviceRetain;   // режим: Manual
    stCfg    : ST_PidCfg;         // конфигурация по умолчанию
    xResOk   : BOOL;              // ответ Reset()
END_VAR

(* ---- RetainAutoRestoredOnRestart.method.decl.st ---- *)
// Старт ПЛК с режимом Auto в stRetain: ФБ стартует в Auto (хук в первом вызове), выход — из
// stCmd.rManualOut_pct (42 %), интегратор инициализирован шагом инициализации (бит DT_GAP первого
// вызова), дальше регулирование без рывка.
METHOD PRIVATE RetainAutoRestoredOnRestart
VAR
    fbTime   : FB_FakeTime;       // подменное время, старт 1 ч
    fbPid    : FB_PID;            // ФБ под тестом (новый экземпляр = после перезапуска)
    stCmd    : ST_PidCmd;         // команды (GVL_Hmi переживает загрузку как Persistent)
    stRetain : ST_DeviceRetain;   // режим Auto из Persistent Variables
    stCfg    : ST_PidCfg;         // конфигурация теста
    iStep    : INT;               // шаг цикла
    rOutSt   : REAL;              // выход первого вызова
    wStsSt   : WORD;              // wStatus первого вызова
END_VAR

(* ---- RetainAutoRestoredOnRestart.method.impl.st ---- *)
coUnit.TEST('Pid_RetainAuto_RestoredOnRestart');
// источник: tools/reference/pid.py, сценарий retain_auto
stCfg.rKp := 2.0;
stCfg.rTi_s := 10.0;
stRetain.eRemoteMode := E_DeviceMode.Auto;
stCmd.rManualOut_pct := 42.0;
stCmd.rSp_eu := 50.0;
fbPid.rPv_eu := 46.0;                                                                  // e = 4 %
fbPid.xPvValid := TRUE;
fbPid(itfTime := fbTime, stCmd := stCmd, stRetain := stRetain, stCfg := stCfg);       // первый вызов
rOutSt := fbPid.rOut_pct;
wStsSt := fbPid.stSts.stCommon.wStatus;
AssertTrue(Condition := fbPid.Mode = E_DeviceMode.Auto, Message := 'Auto restored from retain');
AssertTrue(Condition := fbPid.Available, Message := 'available in Auto');
FOR iStep := 1 TO 2 DO
    fbTime.Advance(tStep := T#100MS);
    fbPid(itfTime := fbTime, stCmd := stCmd, stRetain := stRetain, stCfg := stCfg);
END_FOR
// ref: retain_auto.out_start
AssertEquals_REAL(Expected := 42.0, Actual := rOutSt, Delta := 1.0E-4, Message := 'output from rManualOut_pct');
AssertEquals_WORD(Expected := GVL_Const.PID_STS_DT_GAP, Actual := wStsSt AND GVL_Const.PID_STS_DT_GAP,
                  Message := 'first call: initialisation step');
// ref: retain_auto.out_2
AssertEquals_REAL(Expected := 42.08, Actual := fbPid.rOut_pct, Delta := 1.0E-4, Message := 'control continues');
coUnit.TEST_FINISHED();

(* ---- SameTimestampNoCalcHoldsOutput.method.decl.st ---- *)
// Второй вызов в тот же момент (dt = 0; P-02): расчёта нет — выход и D прежние, хотя PV
// изменилась; следующий шаг учитывает изменение PV один раз. Расчёт с нулевым шагом дал бы
// всплеск D = Kp·Td/Tf·ΔPV = 10 %.
METHOD PRIVATE SameTimestampNoCalcHoldsOutput
VAR
    fbTime   : FB_FakeTime;       // подменное время, старт 1 ч
    fbPid    : FB_PID;            // ФБ под тестом
    stCmd    : ST_PidCmd;         // команды
    stRetain : ST_DeviceRetain;   // режим
    stCfg    : ST_PidCfg;         // конфигурация теста
    iStep    : INT;               // шаг цикла
    rOutBef  : REAL;              // выход до вызова с тем же временем
    rDBef    : REAL;              // D до него
    rOutSame : REAL;              // выход в вызове с тем же временем
    rDSame   : REAL;              // D в нём
END_VAR

(* ---- SameTimestampNoCalcHoldsOutput.method.impl.st ---- *)
coUnit.TEST('Pid_SameTimestamp_NoCalc_HoldsOutput');
// источник: tools/reference/pid.py, сценарий dt_zero
stCfg.rKp := 1.0;
stCfg.rTi_s := 10.0;
stCfg.rTd_s := 2.0;                                                                    // N = 10: Tf = 0,2 с
stCmd.rManualOut_pct := 40.0;
stCmd.rSp_eu := 50.0;
fbPid.rPv_eu := 50.0;
fbPid.xPvValid := TRUE;
fbPid(itfTime := fbTime, stCmd := stCmd, stRetain := stRetain, stCfg := stCfg);       // t0: Manual
fbTime.Advance(tStep := T#100MS);
stCmd.stCommon.xSetAuto := TRUE;
fbPid(itfTime := fbTime, stCmd := stCmd, stRetain := stRetain, stCfg := stCfg);       // Auto
FOR iStep := 1 TO 5 DO
    fbTime.Advance(tStep := T#100MS);
    fbPid(itfTime := fbTime, stCmd := stCmd, stRetain := stRetain, stCfg := stCfg);
END_FOR
rOutBef := fbPid.rOut_pct;
rDBef := fbPid.stSts.rD_pct;
fbPid.rPv_eu := 49.0;
fbPid(itfTime := fbTime, stCmd := stCmd, stRetain := stRetain, stCfg := stCfg);       // то же время
rOutSame := fbPid.rOut_pct;
rDSame := fbPid.stSts.rD_pct;
fbTime.Advance(tStep := T#100MS);
fbPid(itfTime := fbTime, stCmd := stCmd, stRetain := stRetain, stCfg := stCfg);
// ref: dt_zero.out_before
AssertEquals_REAL(Expected := 40.0, Actual := rOutBef, Delta := 1.0E-4, Message := 'steady output');
// ref: dt_zero.d_before
AssertEquals_REAL(Expected := 0.0, Actual := rDBef, Delta := 1.0E-4, Message := 'no D at constant PV');
// ref: dt_zero.out_same
AssertEquals_REAL(Expected := 40.0, Actual := rOutSame, Delta := 1.0E-4, Message := 'dt = 0: output held');
// ref: dt_zero.d_same
AssertEquals_REAL(Expected := 0.0, Actual := rDSame, Delta := 1.0E-4, Message := 'dt = 0: no D spike');
// ref: dt_zero.out_next
AssertEquals_REAL(Expected := 47.666668, Actual := fbPid.rOut_pct, Delta := 1.0E-4, Message := 'next step: P + I + D');
// ref: dt_zero.d_next
AssertEquals_REAL(Expected := 6.666667, Actual := fbPid.stSts.rD_pct, Delta := 1.0E-4, Message := 'PV step once');
// ref: dt_zero.dt_ms_next
AssertEquals_REAL(Expected := 100.0, Actual := fbPid.stSts.rDt_ms, Delta := 1.0E-3, Message := 'dt of the next step');
coUnit.TEST_FINISHED();

(* ---- SampleComputesOnlyEveryTSample.method.decl.st ---- *)
// Период расчёта tSample = 100 мс при вызовах раз в 10 мс: за 300 мс выход меняется ровно три
// раза (на расчётах), между ними держится; шаг расчёта в Sts — 100 мс.
METHOD PRIVATE SampleComputesOnlyEveryTSample
VAR
    fbTime    : FB_FakeTime;       // подменное время, старт 1 ч
    fbPid     : FB_PID;            // ФБ под тестом
    stCmd     : ST_PidCmd;         // команды
    stRetain  : ST_DeviceRetain;   // режим: старт в Manual
    stCfg     : ST_PidCfg;         // конфигурация теста
    iStep     : INT;               // шаг цикла
    rPrev     : REAL;              // выход прошлого вызова
    uiChanges : UINT;              // сколько раз выход изменился
END_VAR

(* ---- SampleComputesOnlyEveryTSample.method.impl.st ---- *)
coUnit.TEST('Pid_Sample_ComputesOnlyEveryTSample');
// источник: tools/reference/pid.py, сценарий sample
stCfg.rKp := 2.0;
stCfg.rTi_s := 10.0;
stCfg.tSample := T#100MS;
stCmd.rManualOut_pct := 30.0;
stCmd.rSp_eu := 50.0;
fbPid.rPv_eu := 50.0;
fbPid.xPvValid := TRUE;
fbPid(itfTime := fbTime, stCmd := stCmd, stRetain := stRetain, stCfg := stCfg);       // t0: Manual
FOR iStep := 1 TO 10 DO
    fbTime.Advance(tStep := T#10MS);
    fbPid(itfTime := fbTime, stCmd := stCmd, stRetain := stRetain, stCfg := stCfg);
END_FOR
fbTime.Advance(tStep := T#10MS);
stCmd.stCommon.xSetAuto := TRUE;
fbPid(itfTime := fbTime, stCmd := stCmd, stRetain := stRetain, stCfg := stCfg);       // Auto между расчётами
fbPid.rPv_eu := 46.0;                                                                  // e = 4 %
rPrev := fbPid.rOut_pct;
FOR iStep := 1 TO 30 DO                                                                // 300 мс по 10 мс
    fbTime.Advance(tStep := T#10MS);
    fbPid(itfTime := fbTime, stCmd := stCmd, stRetain := stRetain, stCfg := stCfg);
    IF fbPid.rOut_pct <> rPrev THEN
        uiChanges := uiChanges + 1;
    END_IF
    rPrev := fbPid.rOut_pct;
END_FOR
// ref: sample.changes
AssertEquals_UINT(Expected := 3, Actual := uiChanges, Message := 'output changes only on 3 samples');
// ref: sample.dt_ms
AssertEquals_REAL(Expected := 100.0, Actual := fbPid.stSts.rDt_ms, Delta := 1.0E-3, Message := 'dt = tSample');
// ref: sample.out_end
AssertEquals_REAL(Expected := 38.16, Actual := fbPid.rOut_pct, Delta := 1.0E-4, Message := 'output after 3 samples');
coUnit.TEST_FINISHED();

(* ---- SetAutoWithInvalidPvRejected.method.decl.st ---- *)
// Запрос Auto при негодной PV (бит xSetAuto и RequestMode) отклоняется до ProcessMode:
// RejectedFault, бит снят, режим остаётся Manual, каждая команда даёт +1 к uiCmdSeq.
METHOD PRIVATE SetAutoWithInvalidPvRejected
VAR
    fbTime   : FB_FakeTime;       // подменное время, старт 1 ч
    fbPid    : FB_PID;            // ФБ под тестом
    stCmd    : ST_PidCmd;         // команды
    stRetain : ST_DeviceRetain;   // режим: старт в Manual
    stCfg    : ST_PidCfg;         // конфигурация по умолчанию
    xReqOk   : BOOL;              // ответ RequestMode
END_VAR

(* ---- SetAutoWithOosRequestOneCommand.method.decl.st ---- *)
// Запрос Auto при негодной PV вместе со старшим запросом OutOfService в одном вызове (P-13):
// одна команда — результат старшего (Accepted), uiCmdSeq + 1, оба бита сброшены.
METHOD PRIVATE SetAutoWithOosRequestOneCommand
VAR
    fbTime   : FB_FakeTime;       // подменное время, старт 1 ч
    fbPid    : FB_PID;            // ФБ под тестом
    stCmd    : ST_PidCmd;         // команды
    stRetain : ST_DeviceRetain;   // режим
    stCfg    : ST_PidCfg;         // конфигурация теста
END_VAR

(* ---- SetpointNaNHeldTargetWithinSpLimits.method.decl.st ---- *)
// Неконечное задание держит прежнюю цель, но и она остаётся в пределах задания: задание NaN уже
// в первом вызове (связь со SCADA ещё не поднялась) даёт цель rSpMin_eu, а не 0 вне пределов;
// сужение пределов наладчиком, пока задание неконечно, ограничивает удерживаемую цель.
METHOD PRIVATE SetpointNaNHeldTargetWithinSpLimits
VAR
    fbTime   : FB_FakeTime;       // подменное время, старт 1 ч
    fbPid    : FB_PID;            // ФБ под тестом
    stCmd    : ST_PidCmd;         // команды
    stRetain : ST_DeviceRetain;   // режим: Manual
    stCfg    : ST_PidCfg;         // пределы задания 20…80
    uBits    : U_RealBits;        // источник NaN
    rTgtStart : REAL;             // цель в первом вызове при NaN
    rSpStart  : REAL;             // действующее задание в первом вызове
    rTgtValid : REAL;             // цель при задании 70
    rTgtHeld  : REAL;             // цель при NaN после 70
END_VAR

(* ---- SetpointNaNHoldsTargetWarns.method.decl.st ---- *)
// Неконечное задание (NaN из Modbus или расчёта): цель остаётся прежней, предупреждение
// PID_WRN_SP_INVALID и общий бит DEV_STS_WARNING; конечное задание снимает предупреждение.
METHOD PRIVATE SetpointNaNHoldsTargetWarns
VAR
    fbTime   : FB_FakeTime;       // подменное время, старт 1 ч
    fbPid    : FB_PID;            // ФБ под тестом
    stCmd    : ST_PidCmd;         // команды
    stRetain : ST_DeviceRetain;   // режим: Manual
    stCfg    : ST_PidCfg;         // конфигурация по умолчанию
    uBits    : U_RealBits;        // источник NaN
    rTgtNaN  : REAL;              // цель при NaN
    wWrnNaN  : WORD;              // wWarning при NaN
    wStsNaN  : WORD;              // wStatus при NaN
END_VAR

(* ---- SetpointRampRateLimited.method.decl.st ---- *)
// Рампа задания 2 инж. ед./с: ступень операторского задания 40 -> 60 проходится за 10 с; через
// 5 с действующее задание 50 и бит SP_RAMPING, через 10 с — 60 и бит снят; цель — сразу 60.
METHOD PRIVATE SetpointRampRateLimited
VAR
    fbTime   : FB_FakeTime;       // подменное время, старт 1 ч
    fbPid    : FB_PID;            // ФБ под тестом
    stCmd    : ST_PidCmd;         // команды
    stRetain : ST_DeviceRetain;   // режим: Manual
    stCfg    : ST_PidCfg;         // конфигурация теста
    iStep    : INT;               // шаг цикла
    rSp5     : REAL;              // задание через 5 с
    wSts5    : WORD;              // wStatus через 5 с
    rTgt5    : REAL;              // цель через 5 с
END_VAR

(* ---- SetpointRampRateLimited.method.impl.st ---- *)
coUnit.TEST('Pid_SetpointRamp_RateLimited');
// источник: tools/reference/pid.py, сценарий sp_ramp
stCfg.rSpRate_ups := 2.0;
stCmd.rManualOut_pct := 30.0;
stCmd.rSp_eu := 40.0;
fbPid.rPv_eu := 40.0;
fbPid.xPvValid := TRUE;
fbPid(itfTime := fbTime, stCmd := stCmd, stRetain := stRetain, stCfg := stCfg);       // t0: задание 40 сразу
stCmd.rSp_eu := 60.0;
FOR iStep := 1 TO 50 DO                                                                // 5 с
    fbTime.Advance(tStep := T#100MS);
    fbPid(itfTime := fbTime, stCmd := stCmd, stRetain := stRetain, stCfg := stCfg);
END_FOR
rSp5 := fbPid.stSts.rSp_eu;
wSts5 := fbPid.stSts.stCommon.wStatus;
rTgt5 := fbPid.stSts.rSpTarget_eu;
FOR iStep := 1 TO 50 DO                                                                // ещё 5 с
    fbTime.Advance(tStep := T#100MS);
    fbPid(itfTime := fbTime, stCmd := stCmd, stRetain := stRetain, stCfg := stCfg);
END_FOR
// ref: sp_ramp.sp_5s
AssertEquals_REAL(Expected := 50.0, Actual := rSp5, Delta := 1.0E-4, Message := 'SP = 40 + 2 * 5 after 5 s');
AssertEquals_REAL(Expected := 60.0, Actual := rTgt5, Delta := 0.0, Message := 'target at once');
AssertEquals_WORD(Expected := GVL_Const.PID_STS_SP_RAMPING, Actual := wSts5 AND GVL_Const.PID_STS_SP_RAMPING,
                  Message := 'SP_RAMPING while ramping');
// ref: sp_ramp.sp_10s
AssertEquals_REAL(Expected := 60.0, Actual := fbPid.stSts.rSp_eu, Delta := 1.0E-4, Message := 'SP reached after 10 s');
AssertEquals_WORD(Expected := 0, Actual := fbPid.stSts.stCommon.wStatus AND GVL_Const.PID_STS_SP_RAMPING,
                  Message := 'SP_RAMPING cleared');
coUnit.TEST_FINISHED();

(* ---- SetpointRampResumesAfterPvFailure.method.decl.st ---- *)
// Рампа задания (2 инж. ед./с, 40 -> 60) и недостоверная PV: пока PV негодна, расчёта нет и
// действующее задание стоит (44); возврат PV — шаг инициализации с dt = 0, рампа продолжается с
// 44 (не прыгает к цели 60) и через 1 с даёт 46. Бит SP_RAMPING остаётся, пока задание не у цели.
METHOD PRIVATE SetpointRampResumesAfterPvFailure
VAR
    fbTime    : FB_FakeTime;       // подменное время, старт 1 ч
    fbPid     : FB_PID;            // ФБ под тестом
    stCmd     : ST_PidCmd;         // команды
    stRetain  : ST_DeviceRetain;   // режим: Manual
    stCfg     : ST_PidCfg;         // конфигурация теста
    iStep     : INT;               // шаг цикла
    rSp2      : REAL;              // задание через 2 с
    rSpFail   : REAL;              // задание после 1 с с негодной PV
    rSpResume : REAL;              // задание в вызове возврата PV
    wStsRes   : WORD;              // wStatus в вызове возврата PV
END_VAR

(* ---- SetpointRampResumesAfterPvFailure.method.impl.st ---- *)
coUnit.TEST('Pid_SetpointRamp_ResumesAfterPvFailure');
// источник: tools/reference/pid.py, сценарий sp_ramp_pv_fail
stCfg.rSpRate_ups := 2.0;
stCmd.rManualOut_pct := 30.0;
stCmd.rSp_eu := 40.0;
fbPid.rPv_eu := 40.0;
fbPid.xPvValid := TRUE;
fbPid(itfTime := fbTime, stCmd := stCmd, stRetain := stRetain, stCfg := stCfg);       // t0: задание 40 сразу
stCmd.rSp_eu := 60.0;
FOR iStep := 1 TO 20 DO                                                                // 2 с рампы
    fbTime.Advance(tStep := T#100MS);
    fbPid(itfTime := fbTime, stCmd := stCmd, stRetain := stRetain, stCfg := stCfg);
END_FOR
rSp2 := fbPid.stSts.rSp_eu;
fbPid.xPvValid := FALSE;
FOR iStep := 1 TO 10 DO                                                                // 1 с без PV
    fbTime.Advance(tStep := T#100MS);
    fbPid(itfTime := fbTime, stCmd := stCmd, stRetain := stRetain, stCfg := stCfg);
END_FOR
rSpFail := fbPid.stSts.rSp_eu;
fbPid.xPvValid := TRUE;
fbTime.Advance(tStep := T#100MS);
fbPid(itfTime := fbTime, stCmd := stCmd, stRetain := stRetain, stCfg := stCfg);       // PV вернулась
rSpResume := fbPid.stSts.rSp_eu;
wStsRes := fbPid.stSts.stCommon.wStatus;
FOR iStep := 1 TO 10 DO                                                                // ещё 1 с
    fbTime.Advance(tStep := T#100MS);
    fbPid(itfTime := fbTime, stCmd := stCmd, stRetain := stRetain, stCfg := stCfg);
END_FOR
// ref: sp_ramp_pv_fail.sp_2s
AssertEquals_REAL(Expected := 44.0, Actual := rSp2, Delta := 1.0E-4, Message := 'SP = 40 + 2 * 2 after 2 s');
// ref: sp_ramp_pv_fail.sp_fail
AssertEquals_REAL(Expected := 44.0, Actual := rSpFail, Delta := 1.0E-4, Message := 'ramp stops while PV invalid');
// ref: sp_ramp_pv_fail.sp_resume
AssertEquals_REAL(Expected := 44.0, Actual := rSpResume, Delta := 1.0E-4, Message := 'no jump to target on PV return');
AssertEquals_WORD(Expected := GVL_Const.PID_STS_SP_RAMPING, Actual := wStsRes AND GVL_Const.PID_STS_SP_RAMPING,
                  Message := 'SP_RAMPING on PV return');
// ref: sp_ramp_pv_fail.sp_resume_1s
AssertEquals_REAL(Expected := 46.0, Actual := fbPid.stSts.rSp_eu, Delta := 1.0E-4, Message := 'ramp resumes at 2 eu/s');
coUnit.TEST_FINISHED();

(* ---- SpExternalTracksIntoCmd.method.decl.st ---- *)
// Внешнее задание: цель — rSpExt_eu (в пределах rSpMin_eu…rSpMax_eu), ФБ пишет её в
// stCmd.rSp_eu; после снятия xSpExt операторское задание продолжается с того же значения.
METHOD PRIVATE SpExternalTracksIntoCmd
VAR
    fbTime   : FB_FakeTime;       // подменное время, старт 1 ч
    fbPid    : FB_PID;            // ФБ под тестом
    stCmd    : ST_PidCmd;         // команды
    stRetain : ST_DeviceRetain;   // режим: старт в Manual
    stCfg    : ST_PidCfg;         // конфигурация по умолчанию (задание 0…100)
    rCmdSp1  : REAL;              // stCmd.rSp_eu при внешнем задании 63
    rTgt1    : REAL;              // цель при внешнем задании 63
END_VAR

(* ---- SpTrackPvInvalidPvKeepsLastSetpoint.method.decl.st ---- *)
// Слежение задания за PV в Manual (xSpTrackPv) идёт только за годной PV: при обрыве датчика
// (AI держит 0 и снимает xValid) задание оператора и цель остаются последними годными, иначе после
// возврата в Auto регулятор погнал бы процесс к ложному значению.
METHOD PRIVATE SpTrackPvInvalidPvKeepsLastSetpoint
VAR
    fbTime   : FB_FakeTime;       // подменное время, старт 1 ч
    fbPid    : FB_PID;            // ФБ под тестом
    stCmd    : ST_PidCmd;         // команды
    stRetain : ST_DeviceRetain;   // режим
    stCfg    : ST_PidCfg;         // конфигурация теста
    rCmdSpF  : REAL;              // stCmd.rSp_eu при негодной PV
    rTgtF    : REAL;              // цель при негодной PV
END_VAR
